// TIA Portal project "슈룹터 프로젝트 찐찐찐완" (V19)

(* hardware
DEVICE "HMI_1"  KTP700 Basic PN
   slot 0: "HMI_1"  KTP700 Basic PN  6AV2 123-2GB03-0AX0  17.0.0.0
   slot 1: "HMI_RT_1"  KTP700 Basic PN  6AV2 123-2GB03-0AX0  17.0.0.0
   slot 5: "HMI_1.IE_CP_1"  PROFINET Interface  17.0.0.0
      slot 1: "PROFINET Interface_1"  PROFINET Interface
         slot 1: "Port_1"  Port
DEVICE "S7-1200 station_1"  S7-1200 Station
   slot 0: "Rack_0"  S7-1200 Rack  Rack  V1.0
   slot 1: "PLC_1"  CPU 1215C DC/DC/DC  6ES7 215-1AG40-0XB0  V4.5
*)

// ===== PLC "PLC_1"  CPU 1215C DC/DC/DC =====

VAR_GLOBAL   // PLC tag table "Default tag table"
   "Tag_1" AT %I0.2 : Bool;
END_VAR

DATA_BLOCK "Alarm_DB"   // DB1
{ S7_Optimized_Access := 'FALSE' }
VERSION : 0.1
   VAR
      Error_PW_Popup : Bool;
      Success_PW_Popup : Bool;
      Pick_Mode : Bool;
      Keep_Mode : Bool;
      Error_PW_PB : Bool;
      Err_Keep_PB : Bool;
      Error_Keep : Bool;
      Error_Pick : Bool;
      Error_Pick_PB : Bool;
      PW_Check_Done : Bool;
      Home_PB : Bool;
      H_ScreenNumber : Int;
   END_VAR
BEGIN
END_DATA_BLOCK

DATA_BLOCK "Password"   // DB2
{ S7_Optimized_Access := 'TRUE' }
VERSION : 0.1
   VAR
      Input_Password : Int := 0;
      Backspace_PB : Bool;
      Clear_PB : Bool;
      PW_Num_PB : Array[0..9] of Bool;
      CV_Value : Array[1..4] of Bool;
   END_VAR
BEGIN
END_DATA_BLOCK

DATA_BLOCK "Locker"   // DB3
{ S7_Optimized_Access := 'TRUE' }
VERSION : 0.1
   VAR
      Locker_Status : Array[0..8] of Bool;
      Locker_Password : Array[0..8] of Int;
      Selected_Locker_NO : Int := 0;
      Check_Trigger : Bool;
      Keep_PB : Bool;
      Pick_UP_PB : Bool;
      Current_Back_PB : Bool;
      PW_Back_PB : Bool;
      Locker_PB : Array[1..8] of Bool;
      Target_Room_NO : Array[0..8] of Int;
      Door_Check_PB : Bool;
   END_VAR
BEGIN
   Target_Room_NO[1] := 0;
   Target_Room_NO[2] := 1;
   Target_Room_NO[3] := 2;
   Target_Room_NO[4] := 3;
   Target_Room_NO[5] := 4;
   Target_Room_NO[6] := 5;
END_DATA_BLOCK

DATA_BLOCK "비밀번호_DB"   // DB4
{ S7_Optimized_Access := 'TRUE' }
VERSION : 0.1
// stored: InstanceOfName 비밀번호
"비밀번호"
BEGIN
END_DATA_BLOCK

DATA_BLOCK "MFC"   // DB5
{ S7_Optimized_Access := 'FALSE' }
VERSION : 0.1
   VAR
      MFC_연결 : TCON_IP_v4;
      HoldingRegs : Array[0..8] of Word;
      MFC_Flag : Word;
      SOL : Bool;
      MFC_Server : Word;
      MFC_Server_ON : Bool;
   END_VAR
BEGIN
   MFC_연결.LocalPort := 503;
   MFC_연결.InterfaceId := 64;
   MFC_연결.ID := 1;
   MFC_연결.ConnectionType := 11;
   MFC_연결.RemoteAddress.ADDR[1] := 0;
   MFC_연결.RemoteAddress.ADDR[2] := 0;
   MFC_연결.RemoteAddress.ADDR[3] := 0;
   MFC_연결.RemoteAddress.ADDR[4] := 0;
END_DATA_BLOCK

DATA_BLOCK "Arduino"   // DB7
{ S7_Optimized_Access := 'FALSE' }
VERSION : 0.1
   VAR
      AD_연결 : TCON_IP_v4;
      Motor_Run : Array[0..3] of Word;
      Photo_SS : Bool;
      AD_Server : Word;
      AD_Server_ON : Bool;
   END_VAR
BEGIN
   AD_연결.InterfaceId := 64;
   AD_연결.ID := 2;
   AD_연결.ConnectionType := 11;
   AD_연결.RemoteAddress.ADDR[1] := 192;
   AD_연결.RemoteAddress.ADDR[2] := 168;
   AD_연결.RemoteAddress.ADDR[3] := 0;
   AD_연결.RemoteAddress.ADDR[4] := 50;
   AD_연결.LocalPort := 502;
END_DATA_BLOCK

FUNCTION_BLOCK "비밀번호 설정"   // FB1, LAD
{ S7_Optimized_Access := 'TRUE' }
VERSION : 0.1
   VAR_INPUT
      Keep_PB : Bool;
      Status_Back_PB : Bool;
      PW_Back_PB : Bool;
      Input_Password : Int;
      Check_Trigger : Bool;
      Locker_Status : Bool;
      Selected_NO : Int;
      Error_Keep_PB : Bool;
      Door_Open : Bool;
      Door_Done : Bool;
   END_VAR
   VAR_OUTPUT
      Keep_Mode : Bool;
      Error_Keep : Bool;
      Success_Password : Bool;
      Locker_Password : Int;
      Status_OUT : Bool;
      Done : Bool;
   END_VAR
   VAR
      data : Int;
   END_VAR
   VAR_TEMP   // added for the SCL form of the ladder/FBD networks
      _w1 : Bool;
   END_VAR
BEGIN

REGION Network 1
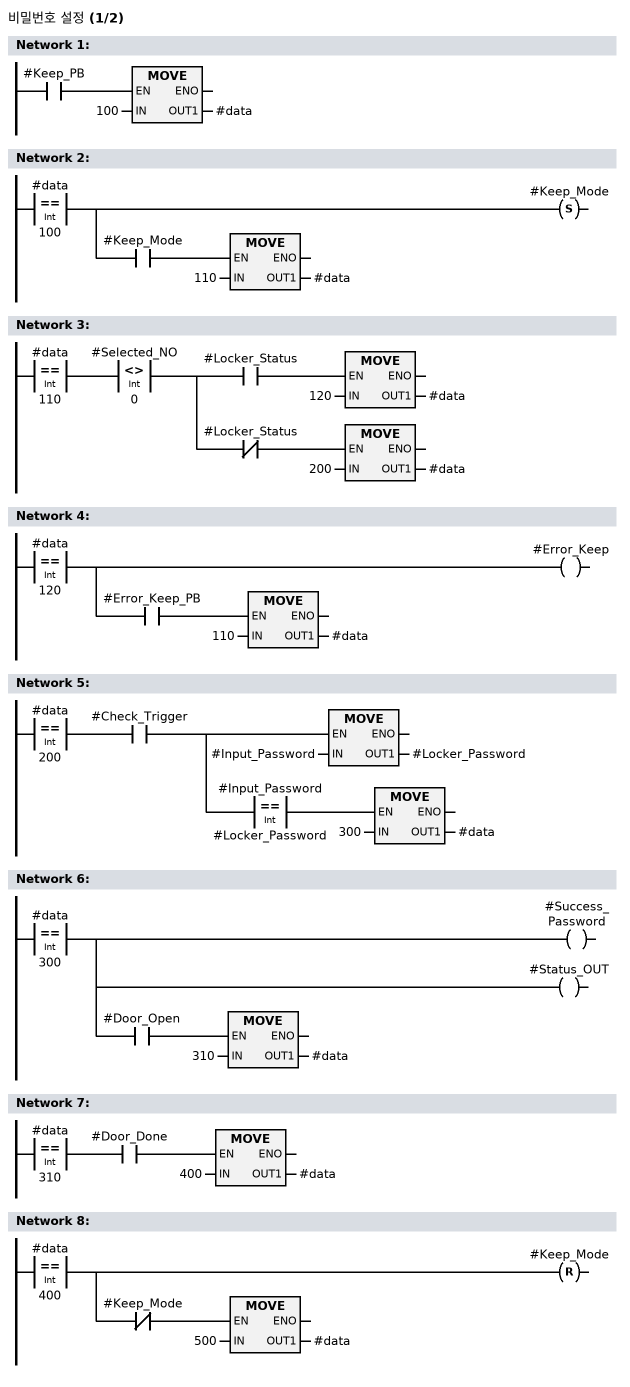
   RUNG wire#powerrail
      Contact( #Keep_PB )
      Move(in := 100, out1 => #data)
   END_RUNG
   // the same network as SCL:
   IF #Keep_PB THEN #data := 100; END_IF;
END_REGION

REGION Network 2
   RUNG wire#powerrail
      { S7_Templates := "SrcType := Int" } EQ_Contact(in1 := #data, in2 := 100)
      wire#w1
      S_Coil( #Keep_Mode )
   END_RUNG
   RUNG wire#w1
      Contact( #Keep_Mode )
      Move(in := 110, out1 => #data)
   END_RUNG
   // the same network as SCL:
   #_w1 := #data = 100;
   IF #_w1 THEN #Keep_Mode := TRUE; END_IF;
   IF #_w1 AND #Keep_Mode THEN #data := 110; END_IF;
END_REGION

REGION Network 3
   RUNG wire#powerrail
      { S7_Templates := "SrcType := Int" } EQ_Contact(in1 := #data, in2 := 110)
      { S7_Templates := "SrcType := Int" } NE_Contact(in1 := #Selected_NO, in2 := 0)
      wire#w1
      Contact( #Locker_Status )
      Move(in := 120, out1 => #data)
   END_RUNG
   RUNG wire#w1
      I_Contact( #Locker_Status )
      Move(in := 200, out1 => #data)
   END_RUNG
   // the same network as SCL:
   #_w1 := (#data = 110) AND (#Selected_NO <> 0);
   IF #_w1 AND #Locker_Status THEN #data := 120; END_IF;
   IF #_w1 AND NOT #Locker_Status THEN #data := 200; END_IF;
END_REGION

REGION Network 4
   RUNG wire#powerrail
      { S7_Templates := "SrcType := Int" } EQ_Contact(in1 := #data, in2 := 120)
      wire#w1
      Coil( #Error_Keep )
   END_RUNG
   RUNG wire#w1
      Contact( #Error_Keep_PB )
      Move(in := 110, out1 => #data)
   END_RUNG
   // the same network as SCL:
   #Error_Keep := #data = 120;
   IF #Error_Keep AND #Error_Keep_PB THEN #data := 110; END_IF;
END_REGION

REGION Network 5
   RUNG wire#powerrail
      { S7_Templates := "SrcType := Int" } EQ_Contact(in1 := #data, in2 := 200)
      Contact( #Check_Trigger )
      wire#w1
      Move(in := #Input_Password, out1 => #Locker_Password)
   END_RUNG
   RUNG wire#w1
      { S7_Templates := "SrcType := Int" } EQ_Contact(in1 := #Input_Password, in2 := #Locker_Password)
      Move(in := 300, out1 => #data)
   END_RUNG
   // the same network as SCL:
   #_w1 := (#data = 200) AND #Check_Trigger;
   IF #_w1 THEN #Locker_Password := #Input_Password; END_IF;
   IF #_w1 AND (#Input_Password = #Locker_Password) THEN #data := 300; END_IF;
END_REGION

REGION Network 6
   RUNG wire#powerrail
      { S7_Templates := "SrcType := Int" } EQ_Contact(in1 := #data, in2 := 300)
      wire#w1
      Coil( #Success_Password )
   END_RUNG
   RUNG wire#w1
      Coil( #Status_OUT )
   END_RUNG
   RUNG wire#w1
      Contact( #Door_Open )
      Move(in := 310, out1 => #data)
   END_RUNG
   // the same network as SCL:
   #Success_Password := #data = 300;
   #Status_OUT := #Success_Password;
   IF #Success_Password AND #Door_Open THEN #data := 310; END_IF;
END_REGION

REGION Network 7
   RUNG wire#powerrail
      { S7_Templates := "SrcType := Int" } EQ_Contact(in1 := #data, in2 := 310)
      Contact( #Door_Done )
      Move(in := 400, out1 => #data)
   END_RUNG
   // the same network as SCL:
   IF (#data = 310) AND #Door_Done THEN #data := 400; END_IF;
END_REGION

REGION Network 8
   RUNG wire#powerrail
      { S7_Templates := "SrcType := Int" } EQ_Contact(in1 := #data, in2 := 400)
      wire#w1
      R_Coil( #Keep_Mode )
   END_RUNG
   RUNG wire#w1
      I_Contact( #Keep_Mode )
      Move(in := 500, out1 => #data)
   END_RUNG
   // the same network as SCL:
   #_w1 := #data = 400;
   IF #_w1 THEN #Keep_Mode := FALSE; END_IF;
   IF #_w1 AND NOT #Keep_Mode THEN #data := 500; END_IF;
END_REGION

REGION Network 9
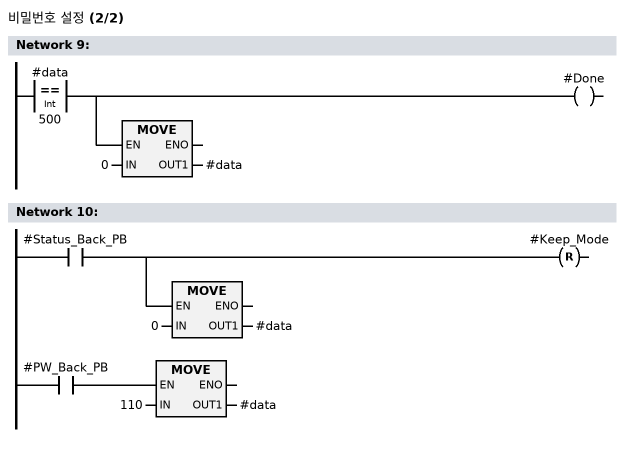
   RUNG wire#powerrail
      { S7_Templates := "SrcType := Int" } EQ_Contact(in1 := #data, in2 := 500)
      wire#w1
      Coil( #Done )
   END_RUNG
   RUNG wire#w1
      Move(in := 0, out1 => #data)
   END_RUNG
   // the same network as SCL:
   #Done := #data = 500;
   IF #Done THEN #data := 0; END_IF;
END_REGION

REGION Network 10
   RUNG wire#powerrail
      Contact( #Status_Back_PB )
      wire#w1
      R_Coil( #Keep_Mode )
   END_RUNG
   RUNG wire#w1
      Move(in := 0, out1 => #data)
   END_RUNG
   RUNG wire#powerrail
      Contact( #PW_Back_PB )
      Move(in := 110, out1 => #data)
   END_RUNG
   // the same network as SCL:
   IF #Status_Back_PB THEN
       #Keep_Mode := FALSE;
       #data := 0;
   END_IF;
   IF #PW_Back_PB THEN #data := 110; END_IF;
END_REGION
END_FUNCTION_BLOCK

FUNCTION_BLOCK "비밀번호 확인"   // FB2, LAD
{ S7_Optimized_Access := 'TRUE' }
VERSION : 0.1
   VAR_INPUT
      Pick_PB : Bool;
      Status_Back_PB : Bool;
      PW_Back_PB : Bool;
      Home_PB : Bool;
      Locker_Status : Bool;
      Selected_NO : Int;
      Input_Password : Int;
      Locker_Password : Int;
      Check_Trigger : Bool;
      Error_PW_PB : Bool;
      Error_Pick_PB : Bool;
      Door_Open : Bool;
      Door_Done : Bool;
   END_VAR
   VAR_OUTPUT
      Pick_Mode : Bool;
      Error_Pick : Bool;
      Error_PW : Bool;
      PW_Check_Success : Bool;
      Status_OUT : Bool;
      Done : Bool;
   END_VAR
   VAR
      data : Int;
   END_VAR
   VAR_TEMP   // added for the SCL form of the ladder/FBD networks
      _w1 : Bool;
   END_VAR
BEGIN

REGION Network 1
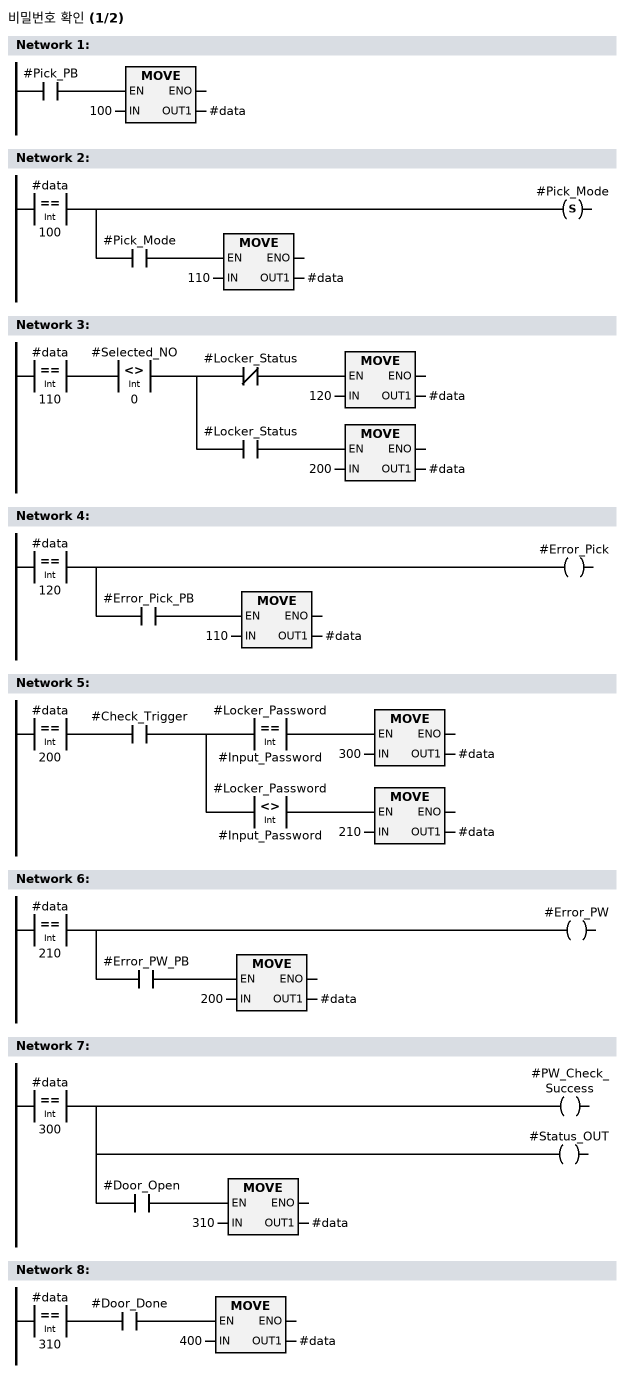
   RUNG wire#powerrail
      Contact( #Pick_PB )
      Move(in := 100, out1 => #data)
   END_RUNG
   // the same network as SCL:
   IF #Pick_PB THEN #data := 100; END_IF;
END_REGION

REGION Network 2
   RUNG wire#powerrail
      { S7_Templates := "SrcType := Int" } EQ_Contact(in1 := #data, in2 := 100)
      wire#w1
      S_Coil( #Pick_Mode )
   END_RUNG
   RUNG wire#w1
      Contact( #Pick_Mode )
      Move(in := 110, out1 => #data)
   END_RUNG
   // the same network as SCL:
   #_w1 := #data = 100;
   IF #_w1 THEN #Pick_Mode := TRUE; END_IF;
   IF #_w1 AND #Pick_Mode THEN #data := 110; END_IF;
END_REGION

REGION Network 3
   RUNG wire#powerrail
      { S7_Templates := "SrcType := Int" } EQ_Contact(in1 := #data, in2 := 110)
      { S7_Templates := "SrcType := Int" } NE_Contact(in1 := #Selected_NO, in2 := 0)
      wire#w1
      I_Contact( #Locker_Status )
      Move(in := 120, out1 => #data)
   END_RUNG
   RUNG wire#w1
      Contact( #Locker_Status )
      Move(in := 200, out1 => #data)
   END_RUNG
   // the same network as SCL:
   #_w1 := (#data = 110) AND (#Selected_NO <> 0);
   IF #_w1 AND NOT #Locker_Status THEN #data := 120; END_IF;
   IF #_w1 AND #Locker_Status THEN #data := 200; END_IF;
END_REGION

REGION Network 4
   RUNG wire#powerrail
      { S7_Templates := "SrcType := Int" } EQ_Contact(in1 := #data, in2 := 120)
      wire#w1
      Coil( #Error_Pick )
   END_RUNG
   RUNG wire#w1
      Contact( #Error_Pick_PB )
      Move(in := 110, out1 => #data)
   END_RUNG
   // the same network as SCL:
   #Error_Pick := #data = 120;
   IF #Error_Pick AND #Error_Pick_PB THEN #data := 110; END_IF;
END_REGION

REGION Network 5
   RUNG wire#powerrail
      { S7_Templates := "SrcType := Int" } EQ_Contact(in1 := #data, in2 := 200)
      Contact( #Check_Trigger )
      wire#w1
      { S7_Templates := "SrcType := Int" } EQ_Contact(in1 := #Locker_Password, in2 := #Input_Password)
      Move(in := 300, out1 => #data)
   END_RUNG
   RUNG wire#w1
      { S7_Templates := "SrcType := Int" } NE_Contact(in1 := #Locker_Password, in2 := #Input_Password)
      Move(in := 210, out1 => #data)
   END_RUNG
   // the same network as SCL:
   #_w1 := (#data = 200) AND #Check_Trigger;
   IF #_w1 AND (#Locker_Password = #Input_Password) THEN #data := 300; END_IF;
   IF #_w1 AND (#Locker_Password <> #Input_Password) THEN #data := 210; END_IF;
END_REGION

REGION Network 6
   RUNG wire#powerrail
      { S7_Templates := "SrcType := Int" } EQ_Contact(in1 := #data, in2 := 210)
      wire#w1
      Coil( #Error_PW )
   END_RUNG
   RUNG wire#w1
      Contact( #Error_PW_PB )
      Move(in := 200, out1 => #data)
   END_RUNG
   // the same network as SCL:
   #Error_PW := #data = 210;
   IF #Error_PW AND #Error_PW_PB THEN #data := 200; END_IF;
END_REGION

REGION Network 7
   RUNG wire#powerrail
      { S7_Templates := "SrcType := Int" } EQ_Contact(in1 := #data, in2 := 300)
      wire#w1
      Coil( #PW_Check_Success )
   END_RUNG
   RUNG wire#w1
      Coil( #Status_OUT )
   END_RUNG
   RUNG wire#w1
      Contact( #Door_Open )
      Move(in := 310, out1 => #data)
   END_RUNG
   // the same network as SCL:
   #PW_Check_Success := #data = 300;
   #Status_OUT := #PW_Check_Success;
   IF #PW_Check_Success AND #Door_Open THEN #data := 310; END_IF;
END_REGION

REGION Network 8
   RUNG wire#powerrail
      { S7_Templates := "SrcType := Int" } EQ_Contact(in1 := #data, in2 := 310)
      Contact( #Door_Done )
      Move(in := 400, out1 => #data)
   END_RUNG
   // the same network as SCL:
   IF (#data = 310) AND #Door_Done THEN #data := 400; END_IF;
END_REGION

REGION Network 9
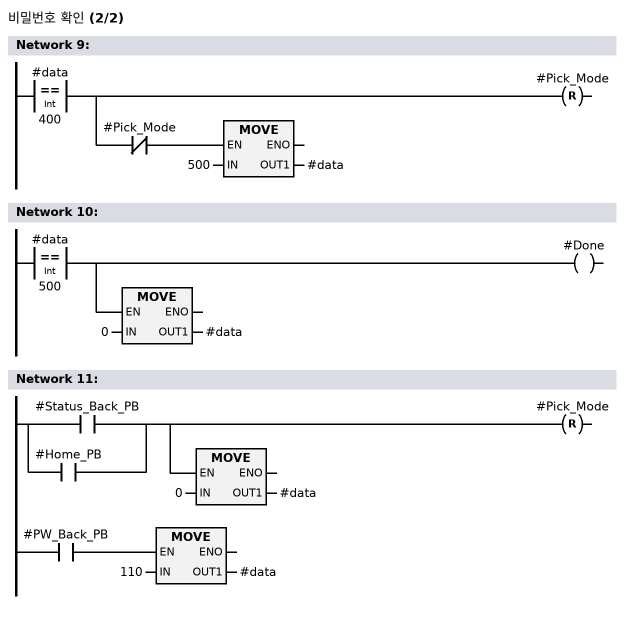
   RUNG wire#powerrail
      { S7_Templates := "SrcType := Int" } EQ_Contact(in1 := #data, in2 := 400)
      wire#w1
      R_Coil( #Pick_Mode )
   END_RUNG
   RUNG wire#w1
      I_Contact( #Pick_Mode )
      Move(in := 500, out1 => #data)
   END_RUNG
   // the same network as SCL:
   #_w1 := #data = 400;
   IF #_w1 THEN #Pick_Mode := FALSE; END_IF;
   IF #_w1 AND NOT #Pick_Mode THEN #data := 500; END_IF;
END_REGION

REGION Network 10
   RUNG wire#powerrail
      { S7_Templates := "SrcType := Int" } EQ_Contact(in1 := #data, in2 := 500)
      wire#w1
      Coil( #Done )
   END_RUNG
   RUNG wire#w1
      Move(in := 0, out1 => #data)
   END_RUNG
   // the same network as SCL:
   #Done := #data = 500;
   IF #Done THEN #data := 0; END_IF;
END_REGION

REGION Network 11
   RUNG wire#powerrail
      Contact( #Status_Back_PB )
      wire#w1
      R_Coil( #Pick_Mode )
   END_RUNG
   RUNG wire#powerrail
      Contact( #Home_PB )
   END_RUNG wire#w1
   RUNG wire#w1
      Move(in := 0, out1 => #data)
   END_RUNG
   RUNG wire#powerrail
      Contact( #PW_Back_PB )
      Move(in := 110, out1 => #data)
   END_RUNG
   // the same network as SCL:
   IF #Status_Back_PB OR #Home_PB THEN
       #Pick_Mode := FALSE;
       #data := 0;
   END_IF;
   IF #PW_Back_PB THEN #data := 110; END_IF;
END_REGION
END_FUNCTION_BLOCK

FUNCTION_BLOCK "비밀번호"   // FB3, LAD
{ S7_Optimized_Access := 'TRUE' }
VERSION : 0.1
   VAR_INPUT
      Target_Room_NO : Array[0..8] of Int;
      회전검출센서 : Bool;
      Door_Check_PB : Bool;
      Keep_PB : Bool;
      Pick_PB : Bool;
      Home_PB : Bool;
      Status_Back_PB : Bool;
      PW_Back_PB : Bool;
      Error_Keep_PB : Bool;
      Error_PW_PB : Bool;
      Error_Pick_PB : Bool;
      Backspace_PB : Bool;
      Clear_PB : Bool;
      MFC_SOL : Bool;
      Check_Trigger : Bool;
      I_Password_Data_PB : Array[0..9] of Bool;
      Locker_PB : Array[1..8] of Bool;
   END_VAR
   VAR_OUTPUT
      Current_Room_NO : Int;
      Selected_NO : Int;
      Current_PW : Int;
      CV_Value : Array[1..4] of Bool;
      Keep_Mode : Bool;
      Pick_Mode : Bool;
      Error_Keep : Bool;
      Error_Pick : Bool;
      Success_Password : Bool;
      Error_PW : Bool;
      PW_Check_Done : Bool;
      SOL_R : Bool;
      HoldingRegs : Array[0..8] of Word;
      Motor_Run : Array[0..3] of Word;
   END_VAR
   VAR_IN_OUT
      Locker_Status : Array[0..8] of Bool;
      Locker_Password : Array[0..8] of Int;
   END_VAR
   VAR
      busy : Array[0..1] of Bool;
      done : Array[0..1] of Bool;
      Status_OUT : Array[0..1] of Bool;
      Password : Int;
      p : Array[0..1] of Bool;
      n : Array[0..4] of Bool;
      사물함번호_Instance : "사물함번호";
      Input_Password : Int;
      PW_Check : Bool;
      Door_Open : Bool;
      Door_Done : Bool;
      "비밀번호 입력 데이터_Instance" : "비밀번호 입력 데이터";
      "비밀번호 설정_Instance" : "비밀번호 설정";
      "비밀번호 확인_Instance" : "비밀번호 확인";
      Go_Target_Instance : "Go_Target";
      Motor_CCW : Bool;
      Motor_CW : Bool;
      T1 : TON_TIME;
   END_VAR
   VAR_TEMP   // added for the SCL form of the ladder/FBD networks
      _w1 : Bool;
      _w2 : Bool;
      _w3 : Bool;
      _w4 : Bool;
      _w5 : Bool;
   END_VAR
BEGIN

REGION Network 1
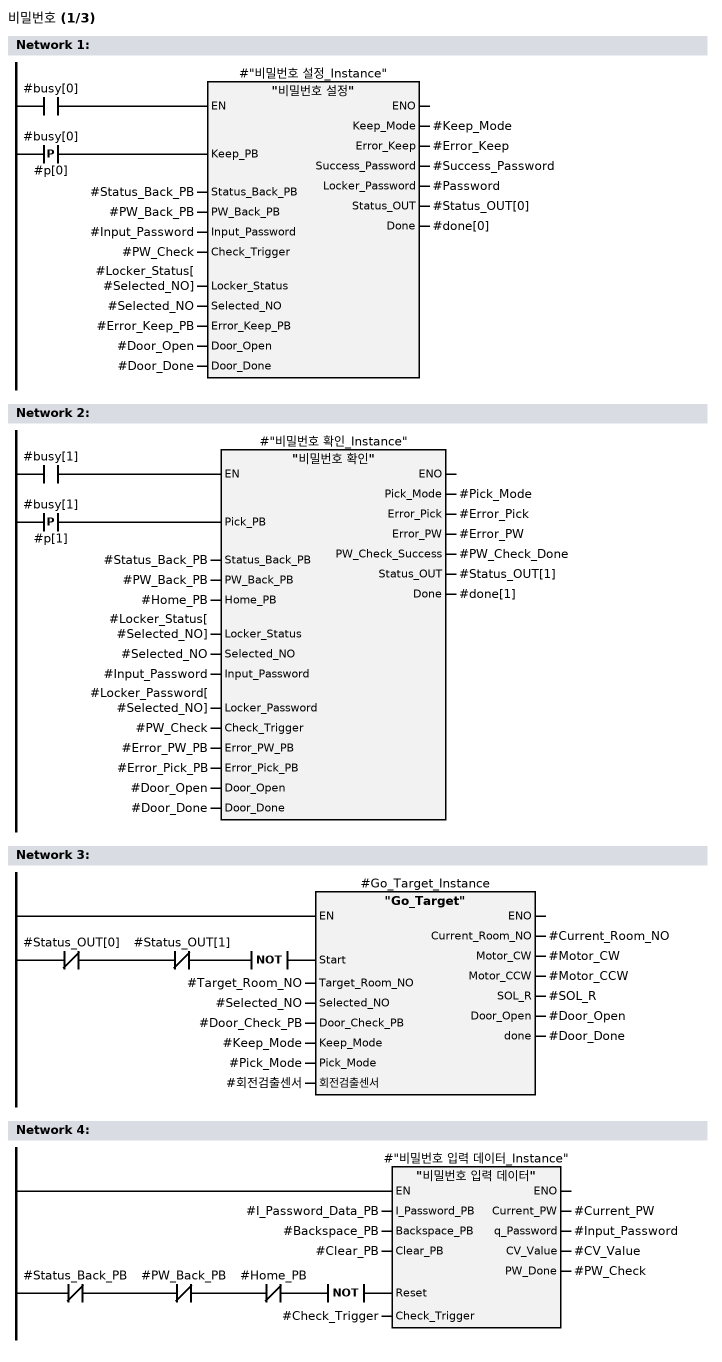
   RUNG wire#powerrail
      Contact( #busy[0] )
      #"비밀번호 설정_Instance"(Keep_PB := wire#w1, Status_Back_PB := #Status_Back_PB, PW_Back_PB := #PW_Back_PB, Input_Password := #Input_Password, Check_Trigger := #PW_Check, Locker_Status := #Locker_Status[#Selected_NO], Selected_NO := #Selected_NO, Error_Keep_PB := #Error_Keep_PB, Door_Open := #Door_Open, Door_Done := #Door_Done, Keep_Mode => #Keep_Mode, Error_Keep => #Error_Keep, Success_Password => #Success_Password, Locker_Password => #Password, Status_OUT => #Status_OUT[0], Done => #done[0])
   END_RUNG
   RUNG wire#powerrail
      P_Contact(operand := #busy[0], bit := #p[0])
   END_RUNG wire#w1
   // the same network as SCL:
   #_w1 := #busy[0] AND NOT #p[0];   // rising edge of #busy[0]
   #p[0] := #busy[0];
   IF #busy[0] THEN
       #"비밀번호 설정_Instance"(Keep_PB := #_w1,   // "비밀번호 설정"
                           Status_Back_PB := #Status_Back_PB,
                           PW_Back_PB := #PW_Back_PB,
                           Input_Password := #Input_Password,
                           Check_Trigger := #PW_Check,
                           Locker_Status := #Locker_Status[#Selected_NO],
                           Selected_NO := #Selected_NO,
                           Error_Keep_PB := #Error_Keep_PB,
                           Door_Open := #Door_Open,
                           Door_Done := #Door_Done,
                           Keep_Mode => #Keep_Mode,
                           Error_Keep => #Error_Keep,
                           Success_Password => #Success_Password,
                           Locker_Password => #Password,
                           Status_OUT => #Status_OUT[0],
                           Done => #done[0]);
   END_IF;
END_REGION

REGION Network 2
   RUNG wire#powerrail
      Contact( #busy[1] )
      #"비밀번호 확인_Instance"(Pick_PB := wire#w1, Status_Back_PB := #Status_Back_PB, PW_Back_PB := #PW_Back_PB, Home_PB := #Home_PB, Locker_Status := #Locker_Status[#Selected_NO], Selected_NO := #Selected_NO, Input_Password := #Input_Password, Locker_Password := #Locker_Password[#Selected_NO], Check_Trigger := #PW_Check, Error_PW_PB := #Error_PW_PB, Error_Pick_PB := #Error_Pick_PB, Door_Open := #Door_Open, Door_Done := #Door_Done, Pick_Mode => #Pick_Mode, Error_Pick => #Error_Pick, Error_PW => #Error_PW, PW_Check_Success => #PW_Check_Done, Status_OUT => #Status_OUT[1], Done => #done[1])
   END_RUNG
   RUNG wire#powerrail
      P_Contact(operand := #busy[1], bit := #p[1])
   END_RUNG wire#w1
   // the same network as SCL:
   #_w1 := #busy[1] AND NOT #p[1];   // rising edge of #busy[1]
   #p[1] := #busy[1];
   IF #busy[1] THEN
       #"비밀번호 확인_Instance"(Pick_PB := #_w1,   // "비밀번호 확인"
                           Status_Back_PB := #Status_Back_PB,
                           PW_Back_PB := #PW_Back_PB,
                           Home_PB := #Home_PB,
                           Locker_Status := #Locker_Status[#Selected_NO],
                           Selected_NO := #Selected_NO,
                           Input_Password := #Input_Password,
                           Locker_Password := #Locker_Password[#Selected_NO],
                           Check_Trigger := #PW_Check,
                           Error_PW_PB := #Error_PW_PB,
                           Error_Pick_PB := #Error_Pick_PB,
                           Door_Open := #Door_Open,
                           Door_Done := #Door_Done,
                           Pick_Mode => #Pick_Mode,
                           Error_Pick => #Error_Pick,
                           Error_PW => #Error_PW,
                           PW_Check_Success => #PW_Check_Done,
                           Status_OUT => #Status_OUT[1],
                           Done => #done[1]);
   END_IF;
END_REGION

REGION Network 3
   RUNG wire#powerrail
      #Go_Target_Instance(Start := wire#w1, Target_Room_NO := #Target_Room_NO, Selected_NO := #Selected_NO, Door_Check_PB := #Door_Check_PB, Keep_Mode := #Keep_Mode, Pick_Mode := #Pick_Mode, 회전검출센서 := #회전검출센서, Current_Room_NO => #Current_Room_NO, Motor_CW => #Motor_CW, Motor_CCW => #Motor_CCW, SOL_R => #SOL_R, Door_Open => #Door_Open, done => #Door_Done)
   END_RUNG
   RUNG wire#powerrail
      I_Contact( #Status_OUT[0] )
      I_Contact( #Status_OUT[1] )
      Not()
   END_RUNG wire#w1
   // the same network as SCL:
   #Go_Target_Instance(Start := NOT (NOT #Status_OUT[0] AND NOT #Status_OUT[1]),   // "Go_Target"
                       Target_Room_NO := #Target_Room_NO,
                       Selected_NO := #Selected_NO,
                       Door_Check_PB := #Door_Check_PB,
                       Keep_Mode := #Keep_Mode,
                       Pick_Mode := #Pick_Mode,
                       회전검출센서 := #회전검출센서,
                       Current_Room_NO => #Current_Room_NO,
                       Motor_CW => #Motor_CW,
                       Motor_CCW => #Motor_CCW,
                       SOL_R => #SOL_R,
                       Door_Open => #Door_Open,
                       done => #Door_Done);
END_REGION

REGION Network 4
   RUNG wire#powerrail
      #"비밀번호 입력 데이터_Instance"(Reset := wire#w1, I_Password_PB := #I_Password_Data_PB, Backspace_PB := #Backspace_PB, Clear_PB := #Clear_PB, Check_Trigger := #Check_Trigger, Current_PW => #Current_PW, q_Password => #Input_Password, CV_Value => #CV_Value, PW_Done => #PW_Check)
   END_RUNG
   RUNG wire#powerrail
      I_Contact( #Status_Back_PB )
      I_Contact( #PW_Back_PB )
      I_Contact( #Home_PB )
      Not()
   END_RUNG wire#w1
   // the same network as SCL:
   #"비밀번호 입력 데이터_Instance"(I_Password_PB := #I_Password_Data_PB,   // "비밀번호 입력 데이터"
                           Backspace_PB := #Backspace_PB,
                           Clear_PB := #Clear_PB,
                           Reset := NOT (NOT #Status_Back_PB AND NOT #PW_Back_PB AND NOT #Home_PB),
                           Check_Trigger := #Check_Trigger,
                           Current_PW => #Current_PW,
                           q_Password => #Input_Password,
                           CV_Value => #CV_Value,
                           PW_Done => #PW_Check);
END_REGION

REGION Network 5
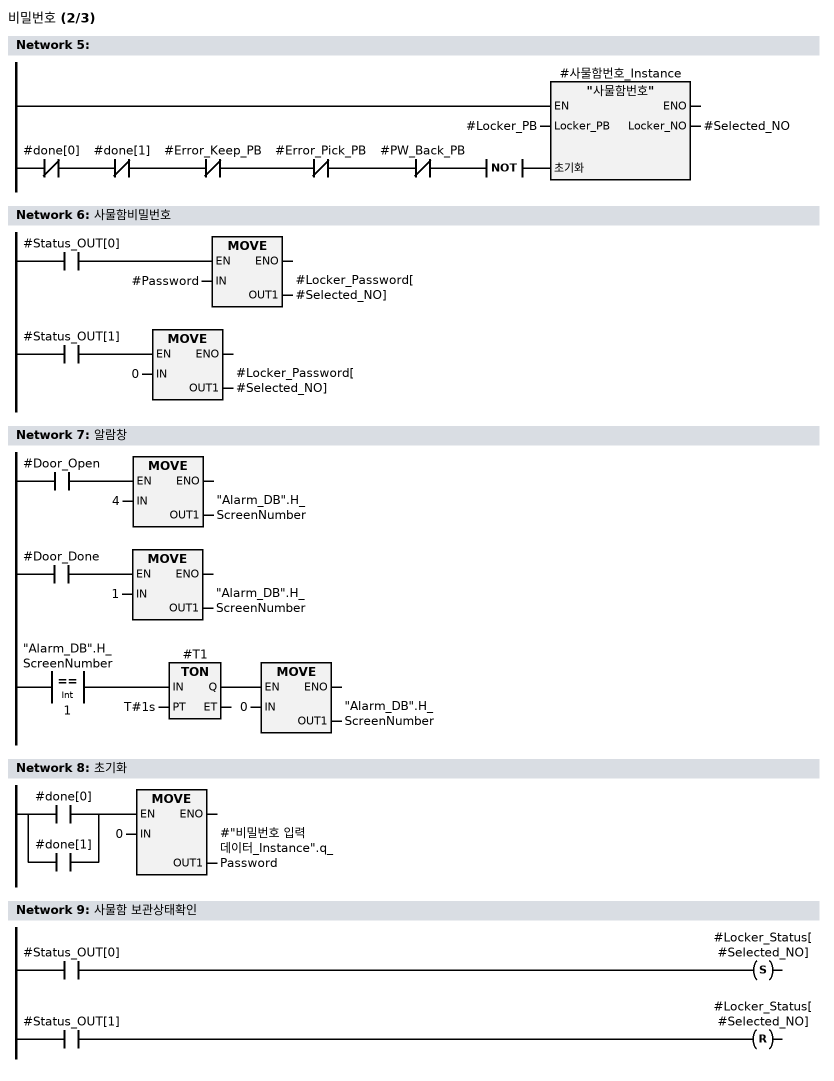
   RUNG wire#powerrail
      #사물함번호_Instance(초기화 := wire#w1, Locker_PB := #Locker_PB, Locker_NO => #Selected_NO)
   END_RUNG
   RUNG wire#powerrail
      I_Contact( #done[0] )
      I_Contact( #done[1] )
      I_Contact( #Error_Keep_PB )
      I_Contact( #Error_Pick_PB )
      I_Contact( #PW_Back_PB )
      Not()
   END_RUNG wire#w1
   // the same network as SCL:
   #사물함번호_Instance(Locker_PB := #Locker_PB,   // "사물함번호"
                   초기화 := NOT (NOT #done[0] AND NOT #done[1] AND NOT #Error_Keep_PB AND NOT #Error_Pick_PB AND NOT #PW_Back_PB),
                   Locker_NO => #Selected_NO);
END_REGION

REGION Network 6: 사물함비밀번호
   RUNG wire#powerrail
      Contact( #Status_OUT[0] )
      Move(in := #Password, out1 => #Locker_Password[#Selected_NO])
   END_RUNG
   RUNG wire#powerrail
      Contact( #Status_OUT[1] )
      Move(in := 0, out1 => #Locker_Password[#Selected_NO])
   END_RUNG
   // the same network as SCL:
   IF #Status_OUT[0] THEN #Locker_Password[#Selected_NO] := #Password; END_IF;
   IF #Status_OUT[1] THEN #Locker_Password[#Selected_NO] := 0; END_IF;
END_REGION

REGION Network 7: 알람창
   IF #Door_Open THEN "Alarm_DB".H_ScreenNumber := 4; END_IF;
   IF #Door_Done THEN "Alarm_DB".H_ScreenNumber := 1; END_IF;
   #T1(IN := "Alarm_DB".H_ScreenNumber = 1, PT := T#1s);   // TON
   IF #T1.Q THEN "Alarm_DB".H_ScreenNumber := 0; END_IF;
END_REGION

REGION Network 8: 초기화
   RUNG wire#powerrail
      Contact( #done[0] )
      wire#w1
      Move(in := 0, out1 => #"비밀번호 입력 데이터_Instance".q_Password)
   END_RUNG
   RUNG wire#powerrail
      Contact( #done[1] )
   END_RUNG wire#w1
   // the same network as SCL:
   IF #done[0] OR #done[1] THEN #"비밀번호 입력 데이터_Instance".q_Password := 0; END_IF;
END_REGION

REGION Network 9: 사물함 보관상태확인
   RUNG wire#powerrail
      Contact( #Status_OUT[0] )
      S_Coil( #Locker_Status[#Selected_NO] )
   END_RUNG
   RUNG wire#powerrail
      Contact( #Status_OUT[1] )
      R_Coil( #Locker_Status[#Selected_NO] )
   END_RUNG
   // the same network as SCL:
   IF #Status_OUT[0] THEN #Locker_Status[#Selected_NO] := TRUE; END_IF;
   IF #Status_OUT[1] THEN #Locker_Status[#Selected_NO] := FALSE; END_IF;
END_REGION

REGION Network 10: 인터록
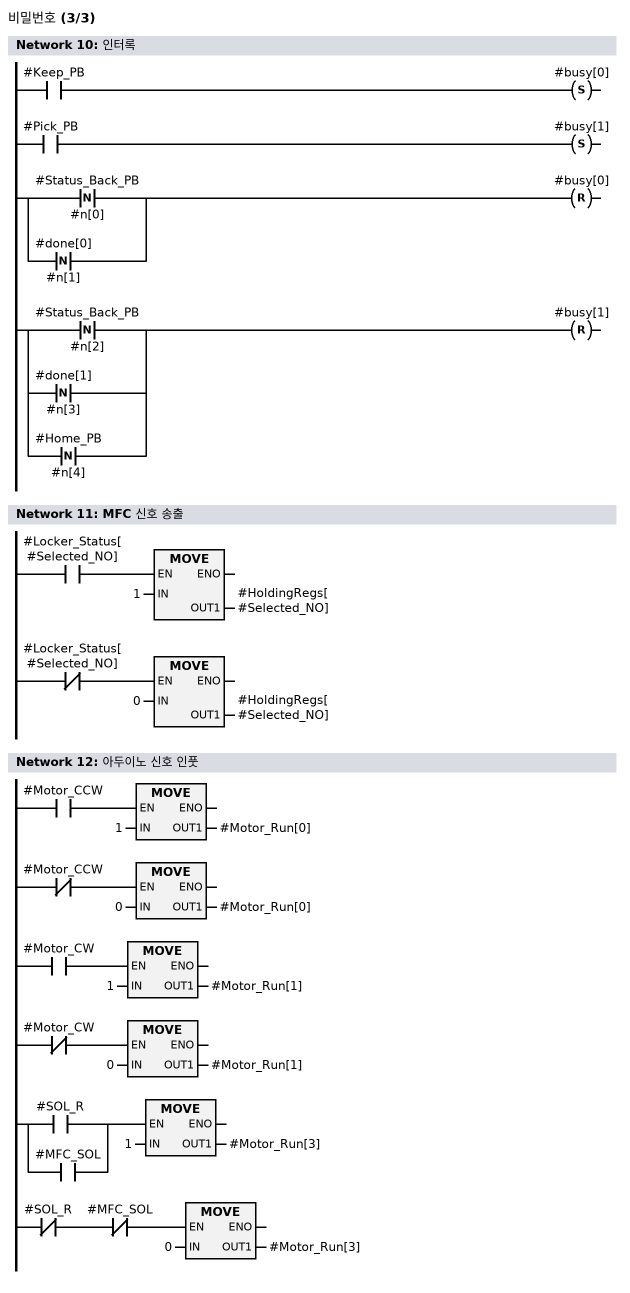
   RUNG wire#powerrail
      Contact( #Keep_PB )
      S_Coil( #busy[0] )
   END_RUNG
   RUNG wire#powerrail
      Contact( #Pick_PB )
      S_Coil( #busy[1] )
   END_RUNG
   RUNG wire#powerrail
      N_Contact(operand := #Status_Back_PB, bit := #n[0])
      wire#w1
      R_Coil( #busy[0] )
   END_RUNG
   RUNG wire#powerrail
      N_Contact(operand := #done[0], bit := #n[1])
   END_RUNG wire#w1
   RUNG wire#powerrail
      N_Contact(operand := #Status_Back_PB, bit := #n[2])
      wire#w2
      R_Coil( #busy[1] )
   END_RUNG
   RUNG wire#powerrail
      N_Contact(operand := #done[1], bit := #n[3])
   END_RUNG wire#w2
   RUNG wire#powerrail
      N_Contact(operand := #Home_PB, bit := #n[4])
   END_RUNG wire#w2
   // the same network as SCL:
   IF #Keep_PB THEN #busy[0] := TRUE; END_IF;
   IF #Pick_PB THEN #busy[1] := TRUE; END_IF;
   #_w1 := NOT #Status_Back_PB AND #n[0];   // falling edge of #Status_Back_PB
   #n[0] := #Status_Back_PB;
   #_w2 := NOT #done[0] AND #n[1];   // falling edge of #done[0]
   #n[1] := #done[0];
   IF #_w1 OR #_w2 THEN #busy[0] := FALSE; END_IF;
   #_w3 := NOT #Status_Back_PB AND #n[2];   // falling edge of #Status_Back_PB
   #n[2] := #Status_Back_PB;
   #_w4 := NOT #done[1] AND #n[3];   // falling edge of #done[1]
   #n[3] := #done[1];
   #_w5 := NOT #Home_PB AND #n[4];   // falling edge of #Home_PB
   #n[4] := #Home_PB;
   IF #_w3 OR #_w4 OR #_w5 THEN #busy[1] := FALSE; END_IF;
END_REGION

REGION Network 11: MFC 신호 송출
   RUNG wire#powerrail
      Contact( #Locker_Status[#Selected_NO] )
      Move(in := 1, out1 => #HoldingRegs[#Selected_NO])
   END_RUNG
   RUNG wire#powerrail
      I_Contact( #Locker_Status[#Selected_NO] )
      Move(in := 0, out1 => #HoldingRegs[#Selected_NO])
   END_RUNG
   // the same network as SCL:
   IF #Locker_Status[#Selected_NO] THEN #HoldingRegs[#Selected_NO] := 1; END_IF;
   IF NOT #Locker_Status[#Selected_NO] THEN #HoldingRegs[#Selected_NO] := 0; END_IF;
END_REGION

REGION Network 12: 아두이노 신호 인풋
   RUNG wire#powerrail
      Contact( #Motor_CCW )
      Move(in := 1, out1 => #Motor_Run[0])
   END_RUNG
   RUNG wire#powerrail
      I_Contact( #Motor_CCW )
      Move(in := 0, out1 => #Motor_Run[0])
   END_RUNG
   RUNG wire#powerrail
      Contact( #Motor_CW )
      Move(in := 1, out1 => #Motor_Run[1])
   END_RUNG
   RUNG wire#powerrail
      I_Contact( #Motor_CW )
      Move(in := 0, out1 => #Motor_Run[1])
   END_RUNG
   RUNG wire#powerrail
      Contact( #SOL_R )
      wire#w1
      Move(in := 1, out1 => #Motor_Run[3])
   END_RUNG
   RUNG wire#powerrail
      Contact( #MFC_SOL )
   END_RUNG wire#w1
   RUNG wire#powerrail
      I_Contact( #SOL_R )
      I_Contact( #MFC_SOL )
      Move(in := 0, out1 => #Motor_Run[3])
   END_RUNG
   // the same network as SCL:
   IF #Motor_CCW THEN #Motor_Run[0] := 1; END_IF;
   IF NOT #Motor_CCW THEN #Motor_Run[0] := 0; END_IF;
   IF #Motor_CW THEN #Motor_Run[1] := 1; END_IF;
   IF NOT #Motor_CW THEN #Motor_Run[1] := 0; END_IF;
   IF #SOL_R OR #MFC_SOL THEN #Motor_Run[3] := 1; END_IF;
   IF NOT #SOL_R AND NOT #MFC_SOL THEN #Motor_Run[3] := 0; END_IF;
END_REGION
END_FUNCTION_BLOCK

FUNCTION_BLOCK "사물함번호"   // FB4, LAD
{ S7_Optimized_Access := 'TRUE' }
VERSION : 0.1
   VAR_INPUT
      Locker_PB : Array[1..8] of Bool;
      초기화 : Bool;
   END_VAR
   VAR_OUTPUT
      Locker_NO : Int;
   END_VAR
BEGIN

REGION Network 1
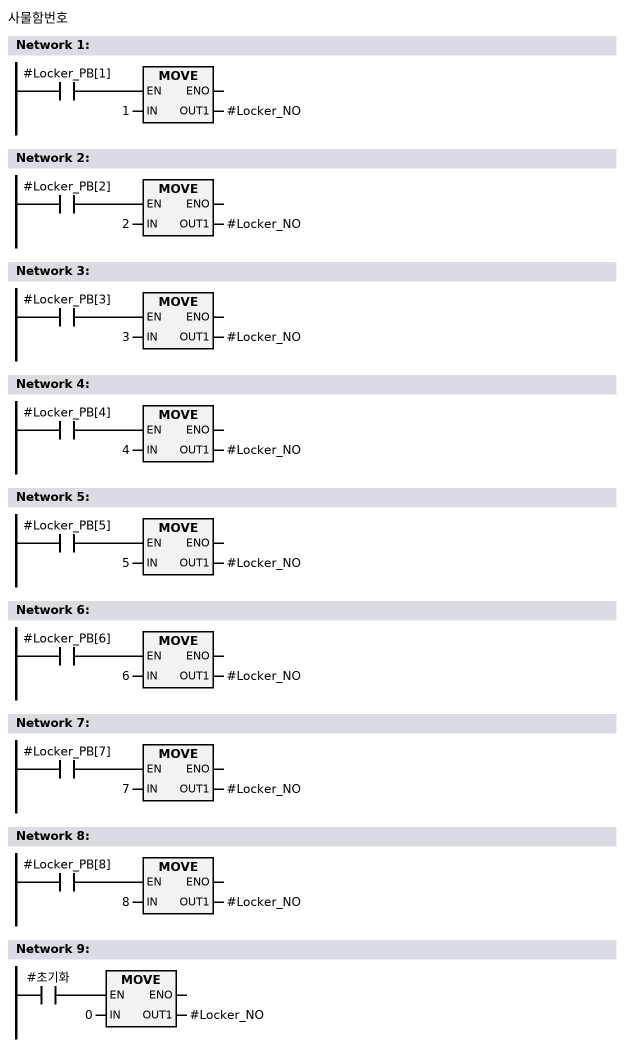
   RUNG wire#powerrail
      Contact( #Locker_PB[1] )
      Move(in := 1, out1 => #Locker_NO)
   END_RUNG
   // the same network as SCL:
   IF #Locker_PB[1] THEN #Locker_NO := 1; END_IF;
END_REGION

REGION Network 2
   RUNG wire#powerrail
      Contact( #Locker_PB[2] )
      Move(in := 2, out1 => #Locker_NO)
   END_RUNG
   // the same network as SCL:
   IF #Locker_PB[2] THEN #Locker_NO := 2; END_IF;
END_REGION

REGION Network 3
   RUNG wire#powerrail
      Contact( #Locker_PB[3] )
      Move(in := 3, out1 => #Locker_NO)
   END_RUNG
   // the same network as SCL:
   IF #Locker_PB[3] THEN #Locker_NO := 3; END_IF;
END_REGION

REGION Network 4
   RUNG wire#powerrail
      Contact( #Locker_PB[4] )
      Move(in := 4, out1 => #Locker_NO)
   END_RUNG
   // the same network as SCL:
   IF #Locker_PB[4] THEN #Locker_NO := 4; END_IF;
END_REGION

REGION Network 5
   RUNG wire#powerrail
      Contact( #Locker_PB[5] )
      Move(in := 5, out1 => #Locker_NO)
   END_RUNG
   // the same network as SCL:
   IF #Locker_PB[5] THEN #Locker_NO := 5; END_IF;
END_REGION

REGION Network 6
   RUNG wire#powerrail
      Contact( #Locker_PB[6] )
      Move(in := 6, out1 => #Locker_NO)
   END_RUNG
   // the same network as SCL:
   IF #Locker_PB[6] THEN #Locker_NO := 6; END_IF;
END_REGION

REGION Network 7
   RUNG wire#powerrail
      Contact( #Locker_PB[7] )
      Move(in := 7, out1 => #Locker_NO)
   END_RUNG
   // the same network as SCL:
   IF #Locker_PB[7] THEN #Locker_NO := 7; END_IF;
END_REGION

REGION Network 8
   RUNG wire#powerrail
      Contact( #Locker_PB[8] )
      Move(in := 8, out1 => #Locker_NO)
   END_RUNG
   // the same network as SCL:
   IF #Locker_PB[8] THEN #Locker_NO := 8; END_IF;
END_REGION

REGION Network 9
   RUNG wire#powerrail
      Contact( #초기화 )
      Move(in := 0, out1 => #Locker_NO)
   END_RUNG
   // the same network as SCL:
   IF #초기화 THEN #Locker_NO := 0; END_IF;
END_REGION
END_FUNCTION_BLOCK

FUNCTION_BLOCK "비밀번호 입력 데이터"   // FB5, LAD
{ S7_Optimized_Access := 'TRUE' }
VERSION : 0.1
   VAR_INPUT
      I_Password_PB : Array[0..9] of Bool;
      Backspace_PB : Bool;
      Clear_PB : Bool;
      Reset : Bool;
      Check_Trigger : Bool;
   END_VAR
   VAR_OUTPUT
      Current_PW : Int;
      q_Password : Int;
      CV_Value : Array[1..4] of Bool;
      PW_Done : Bool;
   END_VAR
   VAR
      PW_data : Int;
      PW_PB_Set_Instance : "PW_PB_Set";
      Start : Bool;
      p : Array[0..2] of Bool;
   END_VAR
   VAR RETAIN
      CTU : CTU_INT;
      data : Int;
   END_VAR
   VAR_TEMP   // added for the SCL form of the ladder/FBD networks
      _w1 : Bool;
      _w2 : Bool;
      _w3 : Bool;
   END_VAR
BEGIN

REGION Network 1
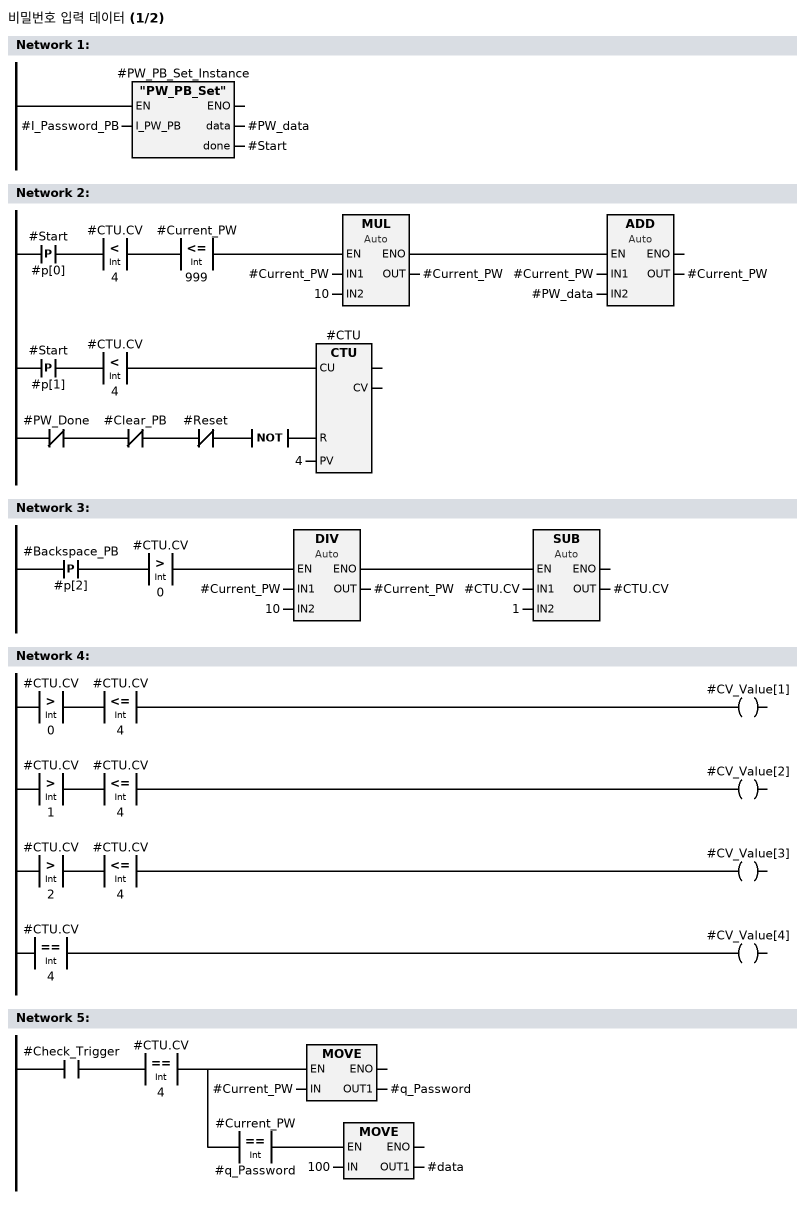
   RUNG wire#powerrail
      #PW_PB_Set_Instance(I_PW_PB := #I_Password_PB, data => #PW_data, done => #Start)
   END_RUNG
   // the same network as SCL:
   #PW_PB_Set_Instance(I_PW_PB := #I_Password_PB, data => #PW_data, done => #Start);   // "PW_PB_Set"
END_REGION

REGION Network 2
   #_w1 := #Start AND NOT #p[0];   // rising edge of #Start
   #p[0] := #Start;
   #_w2 := #_w1 AND (#CTU.CV < 4) AND (#Current_PW <= 999);
   IF #_w2 THEN
       #Current_PW := #Current_PW * 10;
       #Current_PW := #Current_PW + #PW_data;
   END_IF;
   #_w3 := #Start AND NOT #p[1];   // rising edge of #Start
   #p[1] := #Start;
   #CTU(CU := #_w3 AND (#CTU.CV < 4), R := NOT (NOT #PW_Done AND NOT #Clear_PB AND NOT #Reset), PV := 4);   // CTU
END_REGION

REGION Network 3
   RUNG wire#powerrail
      P_Contact(operand := #Backspace_PB, bit := #p[2])
      { S7_Templates := "SrcType := Int" } GT_Contact(in1 := #CTU.CV, in2 := 0)
      Div(in1 := #Current_PW, in2 := 10, out => #Current_PW)
      Sub(in1 := #CTU.CV, in2 := 1, out => #CTU.CV)
   END_RUNG
   // the same network as SCL:
   #_w1 := #Backspace_PB AND NOT #p[2];   // rising edge of #Backspace_PB
   #p[2] := #Backspace_PB;
   IF #_w1 AND (#CTU.CV > 0) THEN
       #Current_PW := #Current_PW / 10;
       #CTU.CV := #CTU.CV - 1;
   END_IF;
END_REGION

REGION Network 4
   RUNG wire#powerrail
      { S7_Templates := "SrcType := Int" } GT_Contact(in1 := #CTU.CV, in2 := 0)
      { S7_Templates := "SrcType := Int" } LE_Contact(in1 := #CTU.CV, in2 := 4)
      Coil( #CV_Value[1] )
   END_RUNG
   RUNG wire#powerrail
      { S7_Templates := "SrcType := Int" } GT_Contact(in1 := #CTU.CV, in2 := 1)
      { S7_Templates := "SrcType := Int" } LE_Contact(in1 := #CTU.CV, in2 := 4)
      Coil( #CV_Value[2] )
   END_RUNG
   RUNG wire#powerrail
      { S7_Templates := "SrcType := Int" } GT_Contact(in1 := #CTU.CV, in2 := 2)
      { S7_Templates := "SrcType := Int" } LE_Contact(in1 := #CTU.CV, in2 := 4)
      Coil( #CV_Value[3] )
   END_RUNG
   RUNG wire#powerrail
      { S7_Templates := "SrcType := Int" } EQ_Contact(in1 := #CTU.CV, in2 := 4)
      Coil( #CV_Value[4] )
   END_RUNG
   // the same network as SCL:
   #CV_Value[1] := (#CTU.CV > 0) AND (#CTU.CV <= 4);
   #CV_Value[2] := (#CTU.CV > 1) AND (#CTU.CV <= 4);
   #CV_Value[3] := (#CTU.CV > 2) AND (#CTU.CV <= 4);
   #CV_Value[4] := #CTU.CV = 4;
END_REGION

REGION Network 5
   RUNG wire#powerrail
      Contact( #Check_Trigger )
      { S7_Templates := "SrcType := Int" } EQ_Contact(in1 := #CTU.CV, in2 := 4)
      wire#w1
      Move(in := #Current_PW, out1 => #q_Password)
   END_RUNG
   RUNG wire#w1
      { S7_Templates := "SrcType := Int" } EQ_Contact(in1 := #Current_PW, in2 := #q_Password)
      Move(in := 100, out1 => #data)
   END_RUNG
   // the same network as SCL:
   #_w1 := #Check_Trigger AND (#CTU.CV = 4);
   IF #_w1 THEN #q_Password := #Current_PW; END_IF;
   IF #_w1 AND (#Current_PW = #q_Password) THEN #data := 100; END_IF;
END_REGION

REGION Network 6
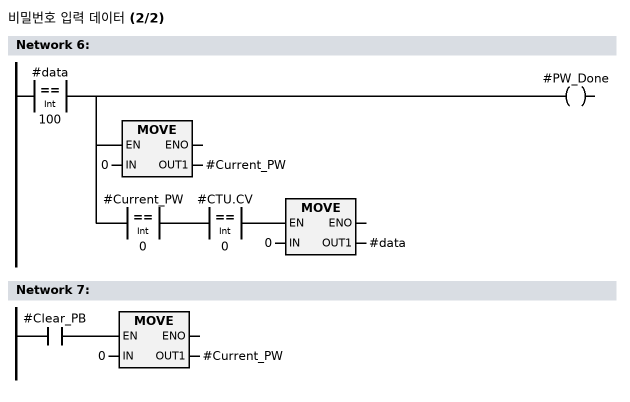
   RUNG wire#powerrail
      { S7_Templates := "SrcType := Int" } EQ_Contact(in1 := #data, in2 := 100)
      wire#w1
      Coil( #PW_Done )
   END_RUNG
   RUNG wire#w1
      Move(in := 0, out1 => #Current_PW)
   END_RUNG
   RUNG wire#w1
      { S7_Templates := "SrcType := Int" } EQ_Contact(in1 := #Current_PW, in2 := 0)
      { S7_Templates := "SrcType := Int" } EQ_Contact(in1 := #CTU.CV, in2 := 0)
      Move(in := 0, out1 => #data)
   END_RUNG
   // the same network as SCL:
   #PW_Done := #data = 100;
   IF #PW_Done THEN #Current_PW := 0; END_IF;
   IF #PW_Done AND (#Current_PW = 0) AND (#CTU.CV = 0) THEN #data := 0; END_IF;
END_REGION

REGION Network 7
   RUNG wire#powerrail
      Contact( #Clear_PB )
      Move(in := 0, out1 => #Current_PW)
   END_RUNG
   // the same network as SCL:
   IF #Clear_PB THEN #Current_PW := 0; END_IF;
END_REGION
END_FUNCTION_BLOCK

FUNCTION_BLOCK "PW_PB_Set"   // FB6, LAD
{ S7_Optimized_Access := 'TRUE' }
VERSION : 0.1
   VAR_INPUT
      I_PW_PB : Array[0..9] of Bool;
   END_VAR
   VAR_OUTPUT
      data : Int;
      done : Bool;
   END_VAR
BEGIN

REGION Network 1
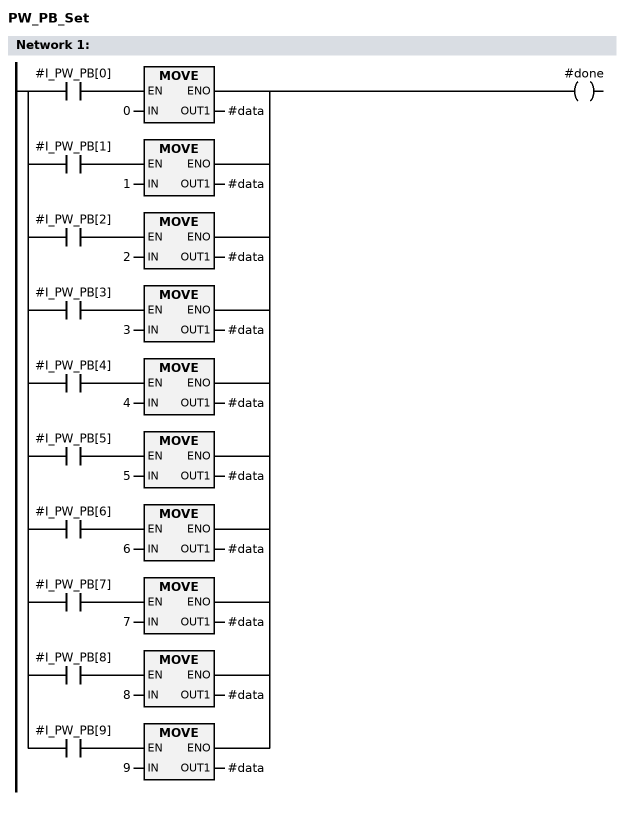
   RUNG wire#powerrail
      Contact( #I_PW_PB[0] )
      Move(in := 0, out1 => #data)
      wire#w1
      Coil( #done )
   END_RUNG
   RUNG wire#powerrail
      Contact( #I_PW_PB[1] )
      Move(in := 1, out1 => #data)
   END_RUNG wire#w1
   RUNG wire#powerrail
      Contact( #I_PW_PB[2] )
      Move(in := 2, out1 => #data)
   END_RUNG wire#w1
   RUNG wire#powerrail
      Contact( #I_PW_PB[3] )
      Move(in := 3, out1 => #data)
   END_RUNG wire#w1
   RUNG wire#powerrail
      Contact( #I_PW_PB[4] )
      Move(in := 4, out1 => #data)
   END_RUNG wire#w1
   RUNG wire#powerrail
      Contact( #I_PW_PB[5] )
      Move(in := 5, out1 => #data)
   END_RUNG wire#w1
   RUNG wire#powerrail
      Contact( #I_PW_PB[6] )
      Move(in := 6, out1 => #data)
   END_RUNG wire#w1
   RUNG wire#powerrail
      Contact( #I_PW_PB[7] )
      Move(in := 7, out1 => #data)
   END_RUNG wire#w1
   RUNG wire#powerrail
      Contact( #I_PW_PB[8] )
      Move(in := 8, out1 => #data)
   END_RUNG wire#w1
   RUNG wire#powerrail
      Contact( #I_PW_PB[9] )
      Move(in := 9, out1 => #data)
   END_RUNG wire#w1
   // the same network as SCL:
   IF #I_PW_PB[0] THEN #data := 0; END_IF;
   IF #I_PW_PB[1] THEN #data := 1; END_IF;
   IF #I_PW_PB[2] THEN #data := 2; END_IF;
   IF #I_PW_PB[3] THEN #data := 3; END_IF;
   IF #I_PW_PB[4] THEN #data := 4; END_IF;
   IF #I_PW_PB[5] THEN #data := 5; END_IF;
   IF #I_PW_PB[6] THEN #data := 6; END_IF;
   IF #I_PW_PB[7] THEN #data := 7; END_IF;
   IF #I_PW_PB[8] THEN #data := 8; END_IF;
   IF #I_PW_PB[9] THEN #data := 9; END_IF;
   #done := #I_PW_PB[0] OR #I_PW_PB[1] OR #I_PW_PB[2] OR #I_PW_PB[3] OR #I_PW_PB[4] OR #I_PW_PB[5] OR #I_PW_PB[6] OR #I_PW_PB[7] OR #I_PW_PB[8] OR #I_PW_PB[9];
END_REGION
END_FUNCTION_BLOCK

FUNCTION_BLOCK "Go_Target"   // FB7, LAD
{ S7_Optimized_Access := 'TRUE' }
VERSION : 0.1
   VAR_INPUT
      Start : Bool;
      Target_Room_NO : Array[0..8] of Int;
      Selected_NO : Int;
      Door_Check_PB : Bool;
      Keep_Mode : Bool;
      Pick_Mode : Bool;
      회전검출센서 : Bool;
   END_VAR
   VAR_OUTPUT
      Current_Room_NO : Int;
      Motor_CW : Bool;
      Motor_CCW : Bool;
      SOL_R : Bool;
      Door_Open : Bool;
      done : Bool;
   END_VAR
   VAR
      data : Int;
   END_VAR
   VAR RETAIN
      CTU1 : CTU_INT;
      CTU2 : CTU_INT;
   END_VAR
   VAR
      P : Array[0..1] of Bool;
      q : Array[0..1] of Bool;
      Target_Val : Int;
      Current_Room_Val : Int;
      Keep_Fin : Bool;
      Pick_Fin : Bool;
      T1 : TON_TIME;
      T2 : TON_TIME;
   END_VAR
   VAR_TEMP   // added for the SCL form of the ladder/FBD networks
      _w1 : Bool;
      _w2 : Bool;
   END_VAR
BEGIN

REGION Network 1
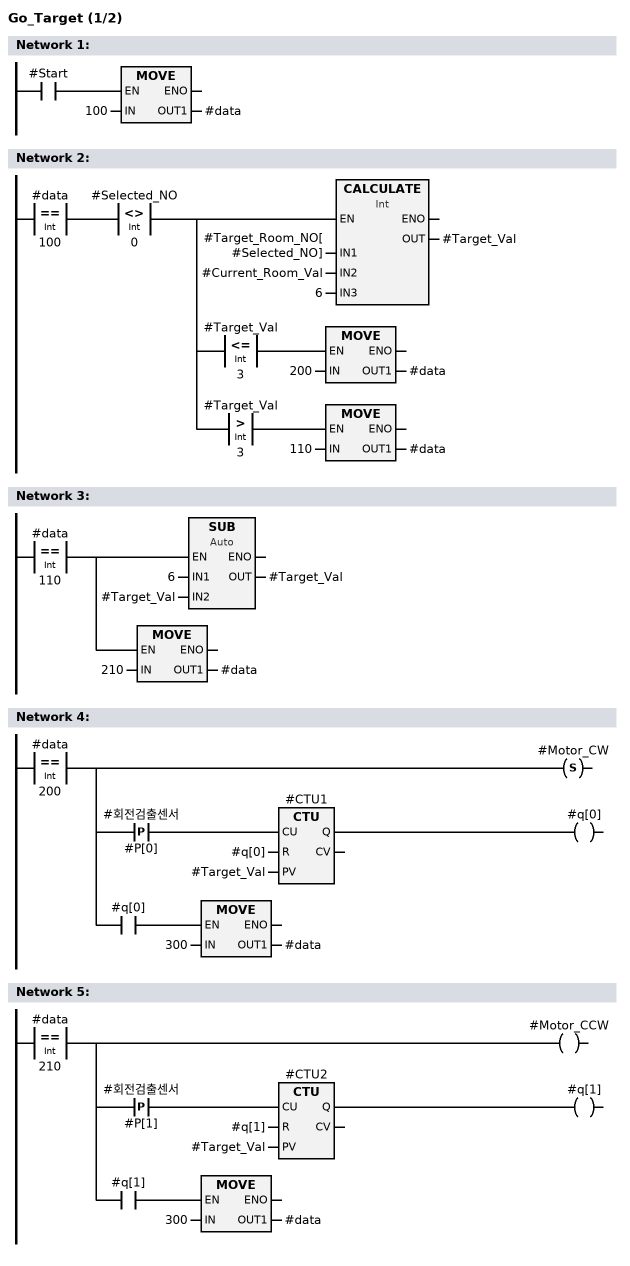
   RUNG wire#powerrail
      Contact( #Start )
      Move(in := 100, out1 => #data)
   END_RUNG
   // the same network as SCL:
   IF #Start THEN #data := 100; END_IF;
END_REGION

REGION Network 2
   RUNG wire#powerrail
      { S7_Templates := "SrcType := Int" } EQ_Contact(in1 := #data, in2 := 100)
      { S7_Templates := "SrcType := Int" } NE_Contact(in1 := #Selected_NO, in2 := 0)
      wire#w1
      { S7_Templates := "SrcType := Int"; S7_Expression := "(IN1 - IN2 + IN3) MOD IN3" } Calculate(in1 := #Target_Room_NO[#Selected_NO], in2 := #Current_Room_Val, in3 := 6, out => #Target_Val)
   END_RUNG
   RUNG wire#w1
      { S7_Templates := "SrcType := Int" } LE_Contact(in1 := #Target_Val, in2 := 3)
      Move(in := 200, out1 => #data)
   END_RUNG
   RUNG wire#w1
      { S7_Templates := "SrcType := Int" } GT_Contact(in1 := #Target_Val, in2 := 3)
      Move(in := 110, out1 => #data)
   END_RUNG
   // the same network as SCL:
   #_w1 := (#data = 100) AND (#Selected_NO <> 0);
   IF #_w1 THEN #Target_Val := (#Target_Room_NO[#Selected_NO] - #Current_Room_Val + 6) MOD 6; END_IF;
   IF #_w1 AND (#Target_Val <= 3) THEN #data := 200; END_IF;
   IF #_w1 AND (#Target_Val > 3) THEN #data := 110; END_IF;
END_REGION

REGION Network 3
   RUNG wire#powerrail
      { S7_Templates := "SrcType := Int" } EQ_Contact(in1 := #data, in2 := 110)
      wire#w1
      Sub(in1 := 6, in2 := #Target_Val, out => #Target_Val)
   END_RUNG
   RUNG wire#w1
      Move(in := 210, out1 => #data)
   END_RUNG
   // the same network as SCL:
   IF #data = 110 THEN
       #Target_Val := 6 - #Target_Val;
       #data := 210;
   END_IF;
END_REGION

REGION Network 4
   #_w1 := #data = 200;
   IF #_w1 THEN #Motor_CW := TRUE; END_IF;
   #_w2 := #_w1 AND #회전검출센서 AND NOT #P[0];   // rising edge of #회전검출센서
   #P[0] := #회전검출센서;
   #CTU1(CU := #_w2, R := #q[0], PV := #Target_Val);   // CTU
   #q[0] := #CTU1.Q;
   IF #_w1 AND #q[0] THEN #data := 300; END_IF;
END_REGION

REGION Network 5
   #Motor_CCW := #data = 210;
   #_w1 := #Motor_CCW AND #회전검출센서 AND NOT #P[1];   // rising edge of #회전검출센서
   #P[1] := #회전검출센서;
   #CTU2(CU := #_w1, R := #q[1], PV := #Target_Val);   // CTU
   #q[1] := #CTU2.Q;
   IF #Motor_CCW AND #q[1] THEN #data := 300; END_IF;
END_REGION

REGION Network 6
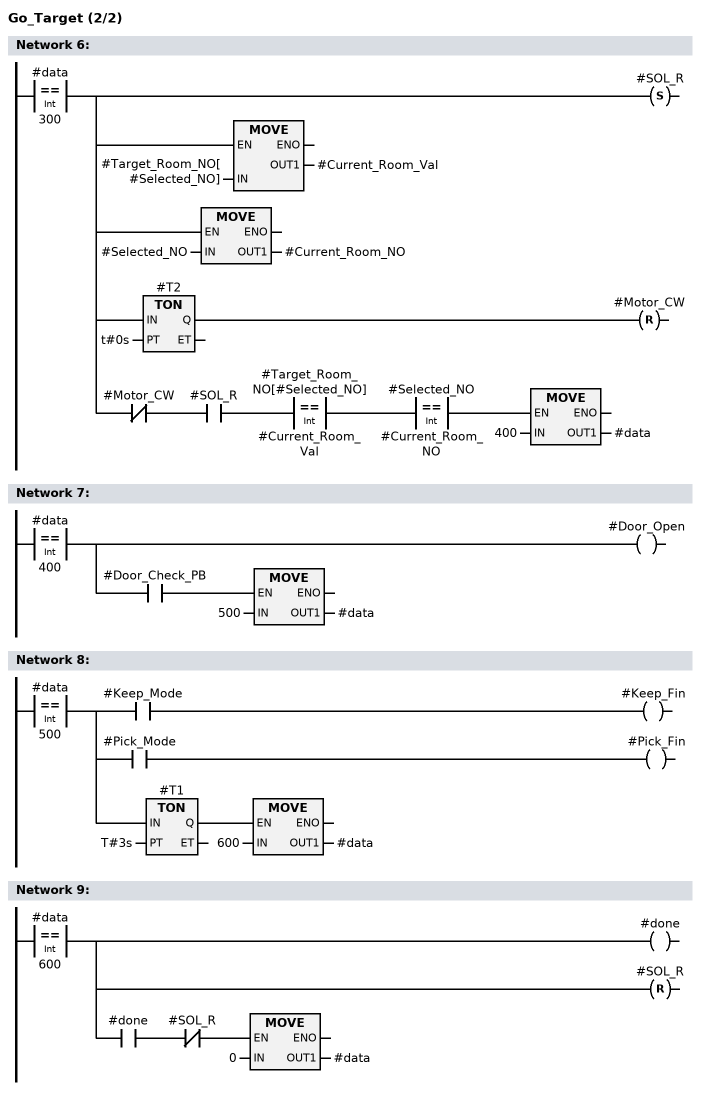
   #_w1 := #data = 300;
   IF #_w1 THEN
       #SOL_R := TRUE;
       #Current_Room_Val := #Target_Room_NO[#Selected_NO];
       #Current_Room_NO := #Selected_NO;
   END_IF;
   #T2(IN := #_w1, PT := t#0s);   // TON
   IF #T2.Q THEN #Motor_CW := FALSE; END_IF;
   IF #_w1 AND NOT #Motor_CW AND #SOL_R AND (#Target_Room_NO[#Selected_NO] = #Current_Room_Val) AND (#Selected_NO = #Current_Room_NO) THEN
       #data := 400;
   END_IF;
END_REGION

REGION Network 7
   RUNG wire#powerrail
      { S7_Templates := "SrcType := Int" } EQ_Contact(in1 := #data, in2 := 400)
      wire#w1
      Coil( #Door_Open )
   END_RUNG
   RUNG wire#w1
      Contact( #Door_Check_PB )
      Move(in := 500, out1 => #data)
   END_RUNG
   // the same network as SCL:
   #Door_Open := #data = 400;
   IF #Door_Open AND #Door_Check_PB THEN #data := 500; END_IF;
END_REGION

REGION Network 8
   #_w1 := #data = 500;
   #Keep_Fin := #_w1 AND #Keep_Mode;
   #Pick_Fin := #_w1 AND #Pick_Mode;
   #T1(IN := #_w1, PT := T#3s);   // TON
   IF #T1.Q THEN #data := 600; END_IF;
END_REGION

REGION Network 9
   RUNG wire#powerrail
      { S7_Templates := "SrcType := Int" } EQ_Contact(in1 := #data, in2 := 600)
      wire#w1
      Coil( #done )
   END_RUNG
   RUNG wire#w1
      R_Coil( #SOL_R )
   END_RUNG
   RUNG wire#w1
      Contact( #done )
      I_Contact( #SOL_R )
      Move(in := 0, out1 => #data)
   END_RUNG
   // the same network as SCL:
   #done := #data = 600;
   IF #done THEN #SOL_R := FALSE; END_IF;
   IF #done AND #done AND NOT #SOL_R THEN #data := 0; END_IF;
END_REGION
END_FUNCTION_BLOCK

FUNCTION_BLOCK "Return_Home"   // FB8, LAD
{ S7_Optimized_Access := 'TRUE' }
VERSION : 0.1
BEGIN
END_FUNCTION_BLOCK

ORGANIZATION_BLOCK "Main"   // OB1, LAD, ProgramCycle
TITLE = "Main Program Sweep (Cycle)"
{ S7_Optimized_Access := 'TRUE' }
VERSION : 0.1
   VAR_INPUT
      Initial_Call : Bool;   // Initial call of this OB
      Remanence : Bool;   // =True, if remanent data are available
   END_VAR
BEGIN

REGION Network 1
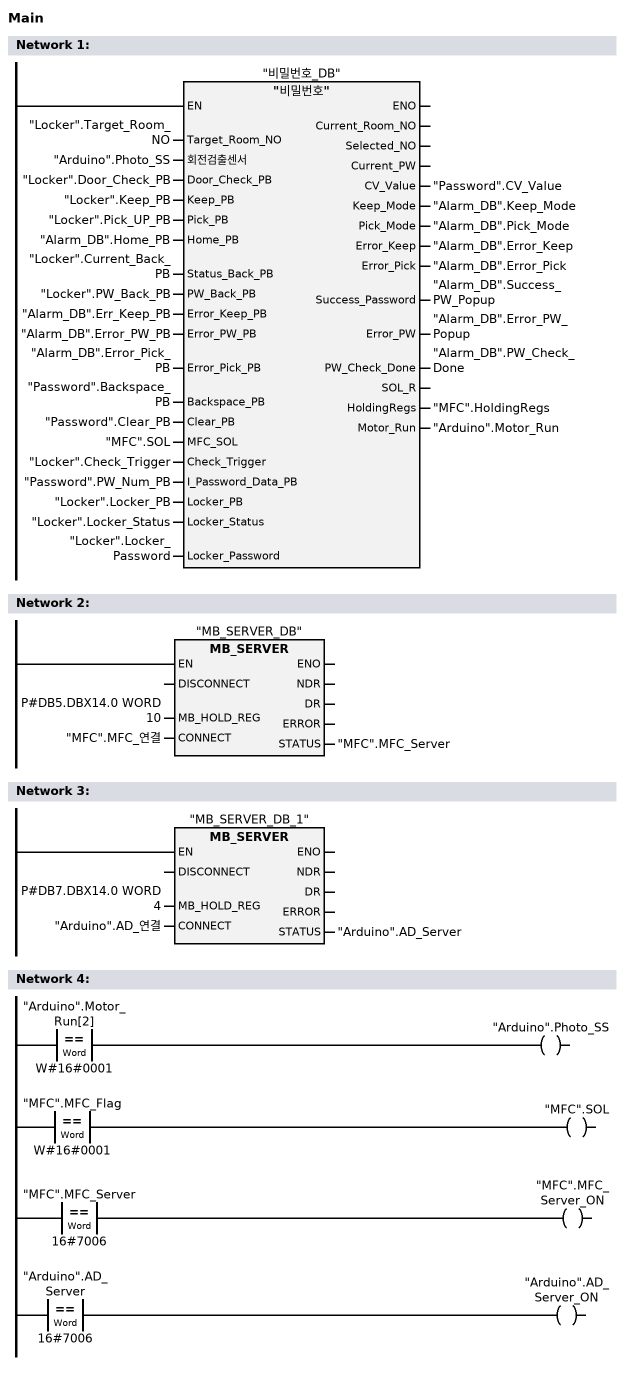
   RUNG wire#powerrail
      "비밀번호_DB"(Target_Room_NO := "Locker".Target_Room_NO, 회전검출센서 := "Arduino".Photo_SS, Door_Check_PB := "Locker".Door_Check_PB, Keep_PB := "Locker".Keep_PB, Pick_PB := "Locker".Pick_UP_PB, Home_PB := "Alarm_DB".Home_PB, Status_Back_PB := "Locker".Current_Back_PB, PW_Back_PB := "Locker".PW_Back_PB, Error_Keep_PB := "Alarm_DB".Err_Keep_PB, Error_PW_PB := "Alarm_DB".Error_PW_PB, Error_Pick_PB := "Alarm_DB".Error_Pick_PB, Backspace_PB := "Password".Backspace_PB, Clear_PB := "Password".Clear_PB, MFC_SOL := "MFC".SOL, Check_Trigger := "Locker".Check_Trigger, I_Password_Data_PB := "Password".PW_Num_PB, Locker_PB := "Locker".Locker_PB, Locker_Status := "Locker".Locker_Status, Locker_Password := "Locker".Locker_Password, Current_Room_NO =>, Selected_NO =>, Current_PW =>, CV_Value => "Password".CV_Value, Keep_Mode => "Alarm_DB".Keep_Mode, Pick_Mode => "Alarm_DB".Pick_Mode, Error_Keep => "Alarm_DB".Error_Keep, Error_Pick => "Alarm_DB".Error_Pick, Success_Password => "Alarm_DB".Success_PW_Popup, Error_PW => "Alarm_DB".Error_PW_Popup, PW_Check_Done => "Alarm_DB".PW_Check_Done, SOL_R =>, HoldingRegs => "MFC".HoldingRegs, Motor_Run => "Arduino".Motor_Run)
   END_RUNG
   // the same network as SCL:
   "비밀번호_DB"(Target_Room_NO := "Locker".Target_Room_NO,   // "비밀번호"
             회전검출센서 := "Arduino".Photo_SS,
             Door_Check_PB := "Locker".Door_Check_PB,
             Keep_PB := "Locker".Keep_PB,
             Pick_PB := "Locker".Pick_UP_PB,
             Home_PB := "Alarm_DB".Home_PB,
             Status_Back_PB := "Locker".Current_Back_PB,
             PW_Back_PB := "Locker".PW_Back_PB,
             Error_Keep_PB := "Alarm_DB".Err_Keep_PB,
             Error_PW_PB := "Alarm_DB".Error_PW_PB,
             Error_Pick_PB := "Alarm_DB".Error_Pick_PB,
             Backspace_PB := "Password".Backspace_PB,
             Clear_PB := "Password".Clear_PB,
             MFC_SOL := "MFC".SOL,
             Check_Trigger := "Locker".Check_Trigger,
             I_Password_Data_PB := "Password".PW_Num_PB,
             Locker_PB := "Locker".Locker_PB,
             Locker_Status := "Locker".Locker_Status,
             Locker_Password := "Locker".Locker_Password,
             CV_Value => "Password".CV_Value,
             Keep_Mode => "Alarm_DB".Keep_Mode,
             Pick_Mode => "Alarm_DB".Pick_Mode,
             Error_Keep => "Alarm_DB".Error_Keep,
             Error_Pick => "Alarm_DB".Error_Pick,
             Success_Password => "Alarm_DB".Success_PW_Popup,
             Error_PW => "Alarm_DB".Error_PW_Popup,
             PW_Check_Done => "Alarm_DB".PW_Check_Done,
             HoldingRegs => "MFC".HoldingRegs,
             Motor_Run => "Arduino".Motor_Run);
END_REGION

REGION Network 2
   "MB_SERVER_DB"(MB_HOLD_REG := P#DB5.DBX14.0 WORD 10, CONNECT := "MFC".MFC_연결, STATUS => "MFC".MFC_Server);   // MB_SERVER
END_REGION

REGION Network 3
   "MB_SERVER_DB_1"(MB_HOLD_REG := P#DB7.DBX14.0 WORD 4,   // MB_SERVER
                    CONNECT := "Arduino".AD_연결,
                    STATUS => "Arduino".AD_Server);
END_REGION

REGION Network 4
   RUNG wire#powerrail
      { S7_Templates := "SrcType := Word" } EQ_Contact(in1 := "Arduino".Motor_Run[2], in2 := W#16#0001)
      Coil( "Arduino".Photo_SS )
   END_RUNG
   RUNG wire#powerrail
      { S7_Templates := "SrcType := Word" } EQ_Contact(in1 := "MFC".MFC_Flag, in2 := W#16#0001)
      Coil( "MFC".SOL )
   END_RUNG
   RUNG wire#powerrail
      { S7_Templates := "SrcType := Word" } EQ_Contact(in1 := "MFC".MFC_Server, in2 := 16#7006)
      Coil( "MFC".MFC_Server_ON )
   END_RUNG
   RUNG wire#powerrail
      { S7_Templates := "SrcType := Word" } EQ_Contact(in1 := "Arduino".AD_Server, in2 := 16#7006)
      Coil( "Arduino".AD_Server_ON )
   END_RUNG
   // the same network as SCL:
   "Arduino".Photo_SS := "Arduino".Motor_Run[2] = W#16#0001;
   "MFC".SOL := "MFC".MFC_Flag = W#16#0001;
   "MFC".MFC_Server_ON := "MFC".MFC_Server = 16#7006;
   "Arduino".AD_Server_ON := "Arduino".AD_Server = 16#7006;
END_REGION
END_ORGANIZATION_BLOCK

(* ===== HMI "HMI_RT_1" =====
system functions are stored by id; their names below are inferred from use
connection "HMI_Connection_1": ETHERNET, SMART_S7_1200_OMS
connection "HMI_Connection_2": ETHERNET, SMART_S7_1200_OMS

HMI tags "Default tag table"
   "Password_Input_Password" : Int = PLC Password.Input_Password, 100 ms
   "Locker_Selected_Locker_NO" : Int = PLC Locker.Selected_Locker_NO, 100 ms
   "Locker_Locker_Status{1}" : Bool = PLC Locker.Locker_Status[1], 100 ms
   "Locker_Locker_Status{2}" : Bool = PLC Locker.Locker_Status[2], 100 ms
   "Locker_Locker_Status{3}" : Bool = PLC Locker.Locker_Status[3], 100 ms
   "Locker_Locker_Status{4}" : Bool = PLC Locker.Locker_Status[4], 100 ms
   "Locker_Locker_Status{5}" : Bool = PLC Locker.Locker_Status[5], 100 ms
   "Locker_Locker_Status{6}" : Bool = PLC Locker.Locker_Status[6], 100 ms
   "Locker_Locker_Status{7}" : Bool = PLC Locker.Locker_Status[7], 100 ms
   "Locker_Locker_Status{8}" : Bool = PLC Locker.Locker_Status[8], 100 ms
   "Locker_Check_Trigger" : Bool = PLC Locker.Check_Trigger, 100 ms
   "Alarm_DB_Error_Password" : Bool = PLC Alarm_DB.Error_PW_Popup AT %DB1.DBX0.0, 100 ms
   "Alarm_DB_Success_Password" : Bool = PLC Alarm_DB.Success_PW_Popup AT %DB1.DBX0.1, 100 ms
   "Tag_ScreenNumber" : Int AT %DB1.DBW0
   "Alarm_DB_Error_PB" : Bool = PLC Alarm_DB.Error_PW_PB AT %DB1.DBX0.4, 100 ms
   "Locker_Keep_PB" : Bool = PLC Locker.Keep_PB, 100 ms
   "Locker_Pick_UP_PB" : Bool = PLC Locker.Pick_UP_PB, 100 ms
   "Alarm_DB_Keep_Mode" : Bool = PLC Alarm_DB.Keep_Mode AT %DB1.DBX0.3, 100 ms
   "Alarm_DB_Pick_Mode" : Bool = PLC Alarm_DB.Pick_Mode AT %DB1.DBX0.2, 100 ms
   "Alarm_DB_Err_Keep_PB" : Bool = PLC Alarm_DB.Err_Keep_PB AT %DB1.DBX0.5, 100 ms
   "Alarm_DB_Error_Keep" : Bool = PLC Alarm_DB.Error_Keep AT %DB1.DBX0.6, 100 ms
   "Alarm_DB_Error_Pick" : Bool = PLC Alarm_DB.Error_Pick AT %DB1.DBX0.7, 100 ms
   "Alarm_DB_Error_Pick_PB" : Bool = PLC Alarm_DB.Error_Pick_PB AT %DB1.DBX1.0, 100 ms
   "Alarm_DB_PW_Check_Done" : Bool = PLC Alarm_DB.PW_Check_Done AT %DB1.DBX1.1, 100 ms
   "Locker_Current_Back_PB" : Bool = PLC Locker.Current_Back_PB, 100 ms
   "Locker_PW_Back_PB" : Bool = PLC Locker.PW_Back_PB, 100 ms
   "Alarm_DB_Home_PB" : Bool = PLC Alarm_DB.Home_PB AT %DB1.DBX1.2, 100 ms
   "Locker_Locker_PB{1}" : Bool = PLC Locker.Locker_PB[1], 100 ms
   "Locker_Locker_PB{2}" : Bool = PLC Locker.Locker_PB[2], 100 ms
   "Locker_Locker_PB{3}" : Bool = PLC Locker.Locker_PB[3], 100 ms
   "Locker_Locker_PB{4}" : Bool = PLC Locker.Locker_PB[4], 100 ms
   "Locker_Locker_PB{5}" : Bool = PLC Locker.Locker_PB[5], 100 ms
   "Locker_Locker_PB{6}" : Bool = PLC Locker.Locker_PB[6], 100 ms
   "Locker_Locker_PB{7}" : Bool = PLC Locker.Locker_PB[7], 100 ms
   "Locker_Locker_PB{8}" : Bool = PLC Locker.Locker_PB[8], 100 ms
   "Password_PW_PB{1}" : Bool = PLC Password.PW_Num_PB[1], 100 ms
   "Password_PW_PB{2}" : Bool = PLC Password.PW_Num_PB[2], 100 ms
   "Password_PW_PB{3}" : Bool = PLC Password.PW_Num_PB[3], 100 ms
   "Password_PW_PB{4}" : Bool = PLC Password.PW_Num_PB[4], 100 ms
   "Password_PW_PB{5}" : Bool = PLC Password.PW_Num_PB[5], 100 ms
   "Password_PW_PB{6}" : Bool = PLC Password.PW_Num_PB[6], 100 ms
   "Password_PW_PB{7}" : Bool = PLC Password.PW_Num_PB[7], 100 ms
   "Password_PW_PB{8}" : Bool = PLC Password.PW_Num_PB[8], 100 ms
   "Password_PW_PB{9}" : Bool = PLC Password.PW_Num_PB[9], 100 ms
   "Password_PW_PB{0}" : Bool = PLC Password.PW_Num_PB[0], 100 ms
   "Password_Backspace_PB" : Bool = PLC Password.Backspace_PB, 100 ms
   "Password_CV_Value{1}" : Bool = PLC Password.CV_Value[1], 100 ms
   "Password_CV_Value{2}" : Bool = PLC Password.CV_Value[2], 100 ms
   "Password_CV_Value{3}" : Bool = PLC Password.CV_Value[3], 100 ms
   "Password_CV_Value{4}" : Bool = PLC Password.CV_Value[4], 100 ms
   "Password_Clear_PB" : Bool = PLC Password.Clear_PB, 100 ms
   "Locker_Door_Check_PB" : Bool = PLC Locker.Door_Check_PB, 100 ms
   "비밀번호_DB_Go_Target_Instance_Keep_Fin" : Bool = PLC 비밀번호_DB.Go_Target_Instance.Keep_Fin, 100 ms
   "비밀번호_DB_Go_Target_Instance_Pick_Fin" : Bool = PLC 비밀번호_DB.Go_Target_Instance.Pick_Fin, 100 ms
   "Alarm_DB_H_ScreenNumber" : Int = PLC Alarm_DB.H_ScreenNumber AT %DB1.DBW2, 100 ms
      on ChangeValue: ActivateScreenByNumber("Alarm_DB_H_ScreenNumber", 0)
   "MFC_MFC_Server_ON" : Bool = PLC MFC.MFC_Server_ON AT %DB5.DBX38.0, 1 s
   "Arduino_AD_Server_ON" : Bool = PLC Arduino.AD_Server_ON AT %DB7.DBX26.0, 1 s

Template "Template_1" 800x480
   Button "Exit" at 714,429 size 71x50; TextOff 'Exit'; PictureOff "ExitRuntime_KTP700_Basic_PN_TR"; PictureOn "ExitRuntime_KTP700_Basic_PN_TR"
      on Release: StopRuntime(0)
   Button "Start screen" at 14,429 size 71x50; TextOff 'Start screen'; PictureOff "NavigateHome_KTP700_Basic_PN_TR"; PictureOn "NavigateHome_KTP700_Basic_PN_TR"
      on Release: ActivateScreen("Root screen", 0)

screen "Root screen" 800x480, template "Template_1"
   Button "HmiScreenItemData" at 25,127 size 355x175; TextOff '보관'; PictureOn "Navigates to Screen0 for KTP700 Basic+ PN 17.0.0.0"; PictureOff "icons8-locker-50"
      on Press: function_b14e0dd5("Locker_Keep_PB", 0)
      on Release: ActivateScreen("Current_Status", 0)
   Button "HmiScreenItemData_1" at 415,127 size 355x175; TextOff '찾기'; PictureOn "Navigates to Screen1 for KTP700 Basic+ PN 17.0.0.0"; PictureOff "icons8-google-web-search-50"
      on Press: function_b14e0dd5("Locker_Pick_UP_PB", 0)
      on Release: ActivateScreen("Current_Status", 0)
   Button "HmiScreenItemData_3" at 105,356 size 170x90; TextOff '대여'; PictureOn "Navigates to Screen0 for KTP700 Basic+ PN 17.0.0.0"; PictureOff "icons8-rent-64"
   Button "HmiScreenItemData_2" at 315,356 size 170x90; TextOff '반납'; PictureOn "Navigates to Screen0 for KTP700 Basic+ PN 17.0.0.0"; PictureOff "icons8-return-48"
   TextField "Text field_1" at 324,35 size 152x62; Text '슈룹터'
   Button "HmiScreenItemData_4" at 525,356 size 170x90; TextOff '구입'; PictureOn "Navigates to Screen0 for KTP700 Basic+ PN 17.0.0.0"; PictureOff "icons8-shop-48"
   TextField "Text field_2" at 148,259 size 119x23; Text '우산 보관 등록'
   TextField "Text field_3" at 554,259 size 119x23; Text '보관 우산 검색'
   GraphicView "Graphic view_1" at 170,151 size 55x50; Picture "icons8-locker-50_1"
   GraphicView "Graphic view_2" at 576,151 size 55x50; Picture "icons8-google-web-search-50_1"
   GraphicView "Graphic view_3" at 380,365 size 40x40; Picture "icons8-return-48_1"
   GraphicView "Graphic view_4" at 167,358 size 50x50; Picture "icons8-rent-64_1"
   GraphicView "Graphic view_5" at 590,364 size 40x40; Picture "icons8-shop-48_1"
   GraphicView "Graphic view_9" at 473,35 size 70x70; Picture "icons8-umbrella-64 (2)"
   Circle "Circle_1" at 46,48 size 12x12
      Appearance <- "MFC_MFC_Server_ON"
   TextField "Text field_4" at 59,42 size 41x23; Text 'MFC'
      Appearance <- "MFC_MFC_Server_ON"
   Circle "Circle_2" at 46,73 size 12x12
      Appearance <- "Arduino_AD_Server_ON"
   TextField "Text field_5" at 59,67 size 69x23; Text 'Arduino'
      Appearance <- "Arduino_AD_Server_ON"

screen "Current_Status" 800x480, template "Template_1"
   Button "Back" at 5,5 size 100x45; TextOff 'Back'
      on Press: function_b14e0dd5("Locker_Current_Back_PB", 0)
      on Release: ActivateScreen("Root screen", 0)
   Button "Button_1" at 89,150 size 115x103; TextOff '1'
      Appearance <- "Locker_Locker_Status{1}"
      on Press: function_b14e0dd5("Locker_Locker_PB{1}", 0)
      on Release: ActivateScreen("Password", 0)
   Button "Button_2" at 90,309 size 115x103; TextOff '5'
      Appearance <- "Locker_Locker_Status{5}"
      on Press: function_b14e0dd5("Locker_Locker_PB{5}", 0)
      on Release: ActivateScreen("Password", 0)
   Button "Button_3" at 262,309 size 115x103; TextOff '6'
      Appearance <- "Locker_Locker_Status{6}"
      on Press: function_b14e0dd5("Locker_Locker_PB{6}", 0)
      on Release: ActivateScreen("Password", 0)
   Button "Button_4" at 434,309 size 115x103; TextOff '7'
   Button "Button_5" at 606,309 size 115x103; TextOff '8'
   Button "Button_6" at 261,150 size 115x103; TextOff '2'
      Appearance <- "Locker_Locker_Status{2}"
      on Press: function_b14e0dd5("Locker_Locker_PB{2}", 0)
      on Release: ActivateScreen("Password", 0)
   Button "Button_7" at 433,150 size 115x103; TextOff '3'
      Appearance <- "Locker_Locker_Status{3}"
      on Press: function_b14e0dd5("Locker_Locker_PB{3}", 0)
      on Release: ActivateScreen("Password", 0)
   Button "Button_8" at 606,150 size 115x103; TextOff '4'
      Appearance <- "Locker_Locker_Status{4}"
      on Press: function_b14e0dd5("Locker_Locker_PB{4}", 0)
      on Release: ActivateScreen("Password", 0)
   Group "Group" at 0,0 size 800x480
   TextField "Text field_2" at 315,25 size 171x43; Text '[찾기모드]'
      Visibility <- "Alarm_DB_Pick_Mode"
   TextField "Text field_1" at 315,25 size 171x43; Text '[보관모드]'
      Visibility <- "Alarm_DB_Keep_Mode"

screen "Password" 800x480
   Button "Back" at 5,5 size 100x45; TextOff 'Back'
      on Press: function_b14e0dd5("Locker_PW_Back_PB", 0)
      on Release: ActivateScreen("Current_Status", 0)
   Button "Button_1" at 122,247 size 90x60; TextOff '1'
      on Press: function_b14e0dd5("Password_PW_PB{1}", 0)
   Button "Button_2" at 270,247 size 90x60; TextOff '2'
      on Press: function_b14e0dd5("Password_PW_PB{2}", 0)
   Button "Button_3" at 405,247 size 90x60; TextOff '3'
      on Press: function_b14e0dd5("Password_PW_PB{3}", 0)
   Button "Button_4" at 122,323 size 90x60; TextOff '4'
      on Press: function_b14e0dd5("Password_PW_PB{4}", 0)
   Button "Button_5" at 270,323 size 90x60; TextOff '5'
      on Press: function_b14e0dd5("Password_PW_PB{5}", 0)
   Button "Button_6" at 405,323 size 90x60; TextOff '6'
      on Press: function_b14e0dd5("Password_PW_PB{6}", 0)
   Button "Button_7" at 122,399 size 90x60; TextOff '7'
      on Press: function_b14e0dd5("Password_PW_PB{7}", 0)
   Button "Button_8" at 270,399 size 90x60; TextOff '8'
      on Press: function_b14e0dd5("Password_PW_PB{8}", 0)
   Button "Button_9" at 405,399 size 90x60; TextOff '9'
      on Press: function_b14e0dd5("Password_PW_PB{9}", 0)
   Button "Button_10" at 546,323 size 90x60; TextOff '0'
      on Press: function_b14e0dd5("Password_PW_PB{0}", 0)
   Button "Button_11" at 675,401 size 90x60; TextOff '확인'
      on Press: function_b14e0dd5("Locker_Check_Trigger", 0)
   Button "Button_12" at 546,247 size 90x60; TextOff '◀'
      on Press: function_b14e0dd5("Password_Backspace_PB", 0)
   TextField "Text field_1" at 149,161 size 36x62; Text '*'
      Visibility <- "Password_CV_Value{1}"
   TextField "Text field_2" at 297,161 size 36x62; Text '*'
      Visibility <- "Password_CV_Value{2}"
   TextField "Text field_3" at 432,161 size 36x62; Text '*'
      Visibility <- "Password_CV_Value{3}"
   TextField "Text field_4" at 573,161 size 36x62; Text '*'
      Visibility <- "Password_CV_Value{4}"
   Button "Button_13" at 546,399 size 90x60; TextOff 'Clear'
      on Press: function_b14e0dd5("Password_Clear_PB", 0)
   TextField "Text field_5" at 144,95 size 513x32; Text '비밀번호 4자리 입력 후 확인버튼을 눌러주세요'
   Rectangle "Rectangle_6" at 120,70 size 560x340
      Visibility <- "Alarm_DB_Error_Password"
   TextField "Text field_6" at 315,105 size 153x62; Text '[오류]'
      Visibility <- "Alarm_DB_Error_Password"
   TextField "Text field_7" at 215,210 size 401x90; Text '비밀번호가 틀렸습니다 다시 입력해주세요'
      Visibility <- "Alarm_DB_Error_Password"
   Button "Button_14" at 570,350 size 90x45; TextOff '다시입력'
      on Press: function_b14e0dd5("Alarm_DB_Error_PB", 0)
      Visibility <- "Alarm_DB_Error_Password"
   Button "Button_15" at 470,350 size 90x45; TextOff '처음으로'
      on Press: function_b14e0dd5("Alarm_DB_Home_PB", 0)
      Visibility <- "Alarm_DB_Error_Password"
      on Release: ActivateScreen("Root screen", 0)
   Rectangle "Rectangle_7" at 120,70 size 560x340
      Visibility <- "Alarm_DB_Error_Pick"
   TextField "Text field_10" at 315,105 size 153x62; Text '[오류]'
      Visibility <- "Alarm_DB_Error_Pick"
   Button "Button_16" at 575,353 size 90x46; TextOff '확인'
      on Press: function_b14e0dd5("Alarm_DB_Error_Pick_PB", 0)
      Visibility <- "Alarm_DB_Error_Pick"
      on Release: ActivateScreen("Current_Status", 0)
   TextField "Text field_11" at 215,210 size 317x82; Text '비어있는 방입니다 다시 선택해주세요'
      Visibility <- "Alarm_DB_Error_Pick"
   Rectangle "Rectangle_8" at 120,70 size 560x340
      Visibility <- "Alarm_DB_Success_Password"
   TextField "Text field_9" at 215,210 size 390x47; Text '잠시만 기다려주세요...'
      Visibility <- "Alarm_DB_Success_Password"
   TextField "Text field_8" at 275,105 size 251x62; Text '[설정완료]'
      Visibility <- "Alarm_DB_Success_Password"
   Rectangle "Rectangle_9" at 120,70 size 560x340
      Visibility <- "Alarm_DB_PW_Check_Done"
   TextField "Text field_13" at 215,210 size 390x47; Text '잠시만 기다려주세요...'
      Visibility <- "Alarm_DB_PW_Check_Done"
   TextField "Text field_12" at 295,105 size 268x62; Text '[확인완료!]'
      Visibility <- "Alarm_DB_PW_Check_Done"
   Rectangle "Rectangle_10" at 120,70 size 560x340
      Visibility <- "Alarm_DB_Error_Keep"
   TextField "Text field_14" at 315,105 size 153x62; Text '[오류]'
      Visibility <- "Alarm_DB_Error_Keep"
   Button "Button_19" at 570,350 size 90x45; TextOff '확인'
      on Press: function_b14e0dd5("Alarm_DB_Err_Keep_PB", 0)
      Visibility <- "Alarm_DB_Error_Keep"
      on Release: ActivateScreen("Current_Status", 0)
   TextField "Text field_15" at 215,210 size 401x90; Text '이미 사용중인 방입니다 다시 선택해주세요'
      Visibility <- "Alarm_DB_Error_Keep"
   Group "Group" at 0,0 size 800x480
   TextField "Text field_16" at 315,25 size 171x43; Text '[보관모드]'
      Visibility <- "Alarm_DB_Keep_Mode"
   TextField "Text field_17" at 315,25 size 171x43; Text '[찾기모드]'
      Visibility <- "Alarm_DB_Pick_Mode"
   Group "Group_1" at 120,70 size 560x340
   Group "Group_3" at 120,70 size 560x340
   Group "Group_2" at 120,70 size 560x340
   Group "Group_4" at 120,70 size 560x340
   Group "Group_5" at 120,70 size 560x340

screen "Locker" 800x480
   TextField "Text field_1" at 32,149 size 739x219; Text '안내에 따라 진행해 주세요 ① 문 열기 ② 우산 보관/찾기 ③ 문 닫기 완료 후 하단의 [확인] 버튼을 눌러주세요'
   Button "Button_1" at 660,390 size 90x60; TextOff '확인'
      on Press: function_b14e0dd5("Locker_Door_Check_PB", 0)
   Rectangle "Rectangle_2" at 120,70 size 560x340
      Visibility <- "비밀번호_DB_Go_Target_Instance_Keep_Fin"
   TextField "Text field_2" at 163,174 size 475x133; Text '우산 보관이 완료되었습니다 이용해주셔서 감사합니다'
      Visibility <- "비밀번호_DB_Go_Target_Instance_Keep_Fin"
   Rectangle "Rectangle_3" at 120,70 size 560x340
      Visibility <- "비밀번호_DB_Go_Target_Instance_Pick_Fin"
   TextField "Text field_3" at 175,174 size 451x133; Text '우산을 수령해주세요 이용해주셔서 감사합니다'
      Visibility <- "비밀번호_DB_Go_Target_Instance_Pick_Fin"
   Group "Group" at 0,0 size 800x480
   TextField "Text field_17" at 315,25 size 171x43; Text '[찾기모드]'
      Visibility <- "Alarm_DB_Pick_Mode"
   TextField "Text field_16" at 315,25 size 171x43; Text '[보관모드]'
      Visibility <- "Alarm_DB_Keep_Mode"
   Group "Group_1" at 120,70 size 560x340
   Group "Group_2" at 120,70 size 560x340
*)